	E_LightTowerState.eRed:;
		qLedGreen	:=FALSE;
		qLedYellow	:=FALSE;
		qLedRed		:=TRUE;
		qLedBlue	:=FALSE;
		IF bBuzzerMuteMemo THEN;
			eBuzzerMode:=eBuzzerOff;
		ELSE
			eBuzzerMode:=eBuzzerError;
		END_IF
		
	E_LightTowerState.eBlue:;
		qLedGreen	:=FALSE;
		qLedYellow	:=FALSE;
		qLedRed		:=FALSE;
		qLedBlue	:=TRUE;
		eBuzzerMode:=eBuzzerOff;	
				
END_CASE


IF qLedRed THEN;
	qSignal_1:=TRUE;	//wire BN
	qSignal_2:=FALSE;	//wire GY
	qSignal_3:=FALSE;	//wire BK
	qSignal_4:=FALSE;	//wire WT	
ELSIF qLedYellow THEN;
	qSignal_1:=TRUE;	//wire BN
	qSignal_2:=FALSE;	//wire GY
	qSignal_3:=FALSE;	//wire BK
	qSignal_4:=TRUE;	//wire WT	
ELSIF qLedGreen THEN;
	qSignal_1:=FALSE;	//wire BN
	qSignal_2:=FALSE;	//wire GY
	qSignal_3:=FALSE;	//wire BK
	qSignal_4:=TRUE;	//wire WT	
ELSIF qLedBlue THEN;
	qSignal_1:=FALSE;	//wire BN
	qSignal_2:=TRUE;	//wire GY
	qSignal_3:=FALSE;	//wire BK
	qSignal_4:=FALSE;	//wire WT	
ELSE;
	qSignal_1:=FALSE;	//wire BN
	qSignal_2:=FALSE;	//wire GY
	qSignal_3:=FALSE;	//wire BK
	qSignal_4:=FALSE;	//wire WT
END_IF
END_METHOD

PROPERTY pState : E_LightTowerState
GET
pState:=eLightTowerState;
END_GET
SET
eLightTowerState:=pState;
END_SET
END_PROPERTY

END_FUNCTION_BLOCK

// ---- 01 Instance/07-Mode/FB_LightTower_Control.TcPOU
FUNCTION_BLOCK FB_LightTower_Control
VAR_INPUT
	ES_State		: BOOL;
	RunProcess1		: BOOL;
	RunProcess2		: BOOL;
	RunProcess3		: BOOL;
	ModeZone1		: E_ModeZone;
	ModeZone2		: E_ModeZone;
	ModeZone3		: E_ModeZone;
END_VAR

VAR_OUTPUT
	eLightTowerState		: E_LightTowerState;
END_VAR
VAR
END_VAR

IF ES_State THEN;
	IF stOper[ModeZone1].iActOperation=E_OperationButtons.ePauseAll 
	OR stOper[ModeZone2].iActOperation=E_OperationButtons.ePauseAll
	OR stOper[ModeZone3].iActOperation=E_OperationButtons.ePauseAll
	THEN;
		eLightTowerState:= E_LightTowerState.eYellow;
	ELSIF RunProcess1 OR RunProcess2 OR RunProcess3 THEN;
		eLightTowerState:= E_LightTowerState.eGreen;
	ELSE;
		eLightTowerState:= E_LightTowerState.eBlue;
	END_IF
	
ELSE;
	eLightTowerState:= E_LightTowerState.eRed;
END_IF

END_FUNCTION_BLOCK

// ---- 03 Project/22 InterConnection/04 Mode/prg_IntCheck.TcPOU
PROGRAM prg_IntCheck
VAR_OUTPUT
	bActive_Marinade_TriB: BOOL;
	bActive_Color_TriB: BOOL;
	bActive_Marinade_Prod: BOOL;
	bActive_Color_Prod: BOOL;
END_VAR

IF fbIntCon_TriB_T1_Marin.bActive OR fbIntCon_TriB_T2_Marin.bActive THEN;
	bActive_Marinade_TriB:=TRUE;
ELSE;
	bActive_Marinade_TriB:=FALSE;
END_IF

IF fbIntCon_TriB_T3_Color.bActive OR fbIntCon_TriB_T4_Color.bActive THEN;
	bActive_Color_TriB:=TRUE;
ELSE;
	bActive_Color_TriB:=FALSE;
END_IF

IF fbIntCon_ProL_T1_Marin.bActive OR fbIntCon_ProL_T2_Marin.bActive THEN;
	bActive_Marinade_Prod:=TRUE;
ELSE;
	bActive_Marinade_Prod:=FALSE;
END_IF

IF fbIntCon_ProL_T3_Color.bActive OR fbIntCon_ProL_T4_Color.bActive THEN;
	bActive_Color_Prod:=TRUE;
ELSE;
	bActive_Color_Prod:=FALSE;
END_IF

END_PROGRAM

// ---- 00 Library/00-General/UserGroup/prg_User.TcPOU
PROGRAM prg_User
VAR
	actUser: E_userGroup:=1;
		
	ton_UserLoged: TON;
	Password: INT;
	ton_Password: TON;
	PT: BOOL;
END_VAR

ton_UserLoged(IN:=actUser<>Group1, PT:=T#10M);

IF ton_UserLoged.Q OR Password=1  THEN
	actUser:=1;
END_IF

IF Password=726 THEN
	actUser:=2;
END_IF

IF Password=345 THEN
	actUser:=3;
END_IF

IF Password=888 THEN
	actUser:=4;
END_IF


ton_Password(IN:=Password<> 0, PT:=T#1s);
IF ton_Password.Q THEN
	Password:=0;
END_IF
;

END_PROGRAM

// ---- 03 Project/22 InterConnection/00 General/prg_InterCon_Usage.TcPOU
PROGRAM prg_InterCon_Usage
VAR
END_VAR

// TriBlender  

IF fbElement[E_Element_List.eTank_1].eState_Short=E_Element_State_Short.eClean 
AND fbElement[E_Element_List.eTriBlender_Marinada].eState_Short=E_Element_State_Short.eClean
THEN;
	//eIntCon_TriB_T1_Marin:=E_InterConnection.Avalable;
END_IF

act_Call_InterConnection();

CASE eTriBlenderUsage OF
	E_TriBlenderUsage.eMarinada_T1,E_TriBlenderUsage.eMarinada_T2:;
		fbElement[E_Element_List.eTriBlender_Marinada].m_StateUpdate_Limit(value:=TRUE);		
		fbElement[E_Element_List.eTriBlender_Color].m_StateUpdate_Limit(value:=TRUE);
	
	E_TriBlenderUsage.eMarinada_Standby:;
		fbElement[E_Element_List.eTriBlender_Marinada].m_StateUpdate_Limit(value:=FALSE);
		fbElement[E_Element_List.eTriBlender_Color].m_StateUpdate_Limit(value:=TRUE);
		
	E_TriBlenderUsage.eColor_T3,E_TriBlenderUsage.eColor_T4:;	
		fbElement[E_Element_List.eTriBlender_Marinada].m_StateUpdate_Limit(value:=TRUE);		
		fbElement[E_Element_List.eTriBlender_Color].m_StateUpdate_Limit(value:=TRUE);
	
	E_TriBlenderUsage.eColor_Standby:;	
		fbElement[E_Element_List.eTriBlender_Marinada].m_StateUpdate_Limit(value:=TRUE);
		fbElement[E_Element_List.eTriBlender_Color].m_StateUpdate_Limit(value:=FALSE);
ELSE;
		fbElement[E_Element_List.eTriBlender_Marinada].m_StateUpdate_Limit(value:=FALSE);
		fbElement[E_Element_List.eTriBlender_Color].m_StateUpdate_Limit(value:=FALSE);	
END_CASE

CASE ePrL_M_Usage OF
	E_PrLine_M_LineUsage.eMarinada_T1,
	E_PrLine_M_LineUsage.eMarinada_T2:;
		fbElement[E_Element_List.eLine_Marinada].m_StateUpdate_Limit(value:=TRUE);
	E_PrLine_M_LineUsage.eNotInUse:;
		fbElement[E_Element_List.eLine_Marinada].m_StateUpdate_Limit(value:=FALSE);
END_CASE

CASE ePrL_C_Usage OF
	E_PrLine_C_Usage.eColor_T3,
	E_PrLine_C_Usage.eColor_T4:;
		fbElement[E_Element_List.eLine_Color].m_StateUpdate_Limit(value:=TRUE);
	E_PrLine_C_Usage.eNotInUse:;
		fbElement[E_Element_List.eLine_Color].m_StateUpdate_Limit(value:=FALSE);
END_CASE
(*
IF eTriBlenderPipe_In=eTriBlenderPipe_Out THEN;
	eTriBlenderPipe:=eTriBlenderPipe_In;
ELSE;
	eTriBlenderPipe:=E_TriBlenderPipe.eNone;
END_IF
*)
(*
CASE fbTriBlender_Select.eStatus OF
	E_TriBlenderSelect.eMarinade:;
		eTriBlenderPipe:=E_TriBlenderPipe.eMarinada;	
	E_TriBlenderSelect.eColor:;
		eTriBlenderPipe:=E_TriBlenderPipe.eColor;
	E_TriBlenderSelect.eDrain:;
		eTriBlenderPipe:=E_TriBlenderPipe.eNone;
ELSE;
	eTriBlenderPipe:=E_TriBlenderPipe.eNone;	
END_CASE
*)

ACTION act_Call_InterConnection:
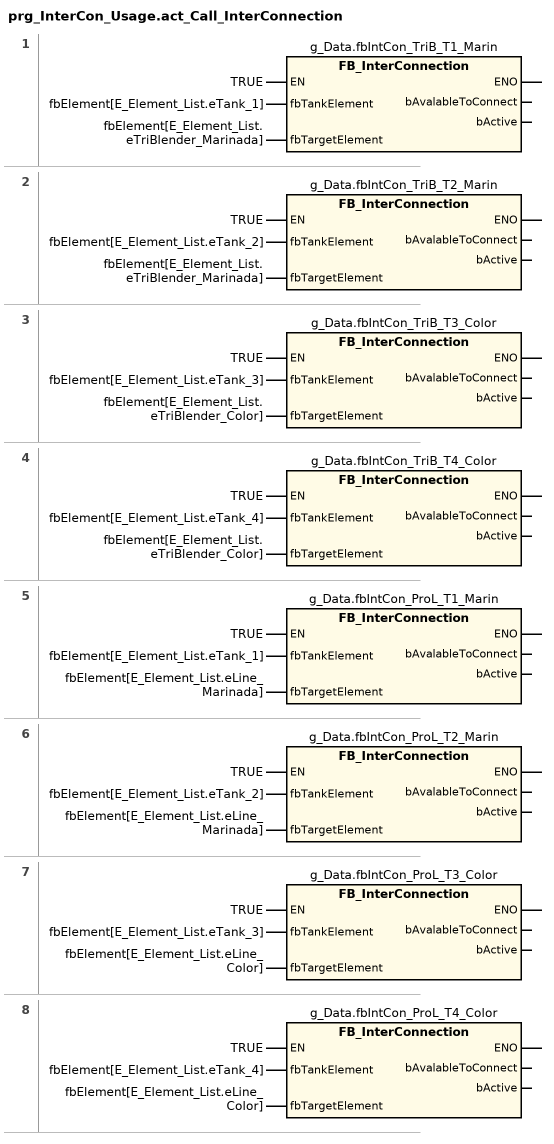
// NETWORK 1
g_Data.fbIntCon_TriB_T1_Marin(fbTankElement := fbElement[E_Element_List.eTank_1], fbTargetElement := fbElement[E_Element_List.eTriBlender_Marinada]); // FB_InterConnection

// NETWORK 2
g_Data.fbIntCon_TriB_T2_Marin(fbTankElement := fbElement[E_Element_List.eTank_2], fbTargetElement := fbElement[E_Element_List.eTriBlender_Marinada]); // FB_InterConnection

// NETWORK 3
g_Data.fbIntCon_TriB_T3_Color(fbTankElement := fbElement[E_Element_List.eTank_3], fbTargetElement := fbElement[E_Element_List.eTriBlender_Color]); // FB_InterConnection

// NETWORK 4
g_Data.fbIntCon_TriB_T4_Color(fbTankElement := fbElement[E_Element_List.eTank_4], fbTargetElement := fbElement[E_Element_List.eTriBlender_Color]); // FB_InterConnection

// NETWORK 5
g_Data.fbIntCon_ProL_T1_Marin(fbTankElement := fbElement[E_Element_List.eTank_1], fbTargetElement := fbElement[E_Element_List.eLine_Marinada]); // FB_InterConnection

// NETWORK 6
g_Data.fbIntCon_ProL_T2_Marin(fbTankElement := fbElement[E_Element_List.eTank_2], fbTargetElement := fbElement[E_Element_List.eLine_Marinada]); // FB_InterConnection

// NETWORK 7
g_Data.fbIntCon_ProL_T3_Color(fbTankElement := fbElement[E_Element_List.eTank_3], fbTargetElement := fbElement[E_Element_List.eLine_Color]); // FB_InterConnection

// NETWORK 8
g_Data.fbIntCon_ProL_T4_Color(fbTankElement := fbElement[E_Element_List.eTank_4], fbTargetElement := fbElement[E_Element_List.eLine_Color]); // FB_InterConnection
END_ACTION

END_PROGRAM

// ---- 03 Project/22 InterConnection/00 General/FB_InterConnection.TcPOU
FUNCTION_BLOCK FB_InterConnection
VAR_INPUT
	//eState_Tank		: E_Element_State_Short;
	//eState_Target	: E_Element_State_Short;
	//eProdType		: E_Product_Type;
	//eTargetTape		: E_Element_Type:=E_Element_Type.eNotSelected;
	reqConnect: BOOL;
	reqDisconnect: BOOL;

END_VAR
VAR_OUTPUT
	bAvalableToConnect: BOOL;
	bAvalableToDisconnect: BOOL;
	bActive: BOOL;
END_VAR
VAR



END_VAR

VAR_IN_OUT
	fbTankElement: FB_Element;
	fbTargetElement: FB_Element;	
END_VAR

act_Avalable();
act_Active();




IF reqConnect THEN;
	m_Connect();
	reqConnect:=FALSE;
END_IF

IF reqDisconnect THEN;
	m_Disconnect();
	reqDisconnect:=FALSE;
END_IF

IF fbTankElement.eInterConnect <> E_InterConnection.NotConnected 
OR fbTargetElement.eInterConnect <> E_InterConnection.NotConnected
THEN;
	m_At_Connected_Pause();
	m_At_Connected_Play();
END_IF

ACTION act_Active:
//fbTargetElement.eState_Long:=fbTankElement.eState_Long;
IF bActive THEN;
	fbTargetElement.m_InterConnected_State(eState_Long_Set:=fbTankElement.eState_Long);
	//fbTargetElement.ExpirationTime:=fbTankElement.ExpirationTime;
	
	CASE fbTargetElement.eType OF		
		E_Element_Type.eLine:;
			//fbTankElement.m_InterConnect(value:=E_InterConnection.ConnToLine);			
		E_Element_Type.eTriBlender:;
			//fbTankElement.m_InterConnect(value:=E_InterConnection.ConnToTriBlender);		
	END_CASE
	//fbTargetElement.m_InterConnect(value:=E_InterConnection.ConnToTank);
	
	CASE fbTankElement.eState_Short OF
		E_Element_State_Short.eNotClean,
		E_Element_State_Short.eClean:;
				//fbTargetElement.ExpirationMode:=E_ExTime.eCIP;

		E_Element_State_Short.eProduct:;
				//fbTargetElement.ExpirationMode:=E_ExTime.eLine;
	END_CASE	

ELSE;
	//fbTankElement.m_Disconnect();
	//fbTargetElement.m_Disconnect();
END_IF
END_ACTION

ACTION act_At_Connected_Pause:

/// Master case
IF fbTankElement.m_Get_Oper_Pause_Puls() THEN;
	CASE fbTankElement.eInterConnect OF 
		E_InterConnection.NotConnected:;
		E_InterConnection.ConnToCIP:;
				// set pause to CIP
				stOper[E_ModeZone.eCIP].bSetPause:=TRUE;
				
		E_InterConnection.ConnToTank:;
				//Not avilble 
		E_InterConnection.ConnToLine:;
				IF fbTargetElement.m_Get_Type()=E_Element_Type.eLine THEN;
					fbTargetElement.m_Set_Oper_Pause();
				END_IF
		E_InterConnection.ConnToTriBlender:;
				IF fbTargetElement.m_Get_Type()=E_Element_Type.eTriBlender THEN;
					fbTargetElement.m_Set_Oper_Pause();
				END_IF				
	END_CASE	
END_IF


/// Slave case
IF fbTargetElement.m_Get_Oper_Pause_Puls() THEN;
	CASE fbTargetElement.eInterConnect OF 
		E_InterConnection.NotConnected:;
		E_InterConnection.ConnToCIP:;
				// set pause to CIP
				stOper[E_ModeZone.eCIP].bSetPause:=TRUE;
				
		E_InterConnection.ConnToTank:;
				IF TRUE
				AND fbTargetElement.m_Get_Type()=E_Element_Type.eLine
				AND fbTankElement.eInterConnect=E_InterConnection.ConnToLine THEN;
					fbTankElement.m_Set_Oper_Pause();
				END_IF
				
				IF TRUE
				AND fbTargetElement.m_Get_Type()=E_Element_Type.eTriBlender
				AND fbTankElement.eInterConnect=E_InterConnection.ConnToTriBlender THEN;
					fbTankElement.m_Set_Oper_Pause();
				END_IF
								
		E_InterConnection.ConnToLine:;
				//Not avilble 
		E_InterConnection.ConnToTriBlender:;
				//Not avilble 			
	END_CASE	
END_IF

// CIP Case
IF stOper[E_ModeZone.eCIP].b_rt_Pause 
AND	fbTankElement.eInterConnect=E_InterConnection.ConnToCIP
THEN;	
	fbTankElement.m_Set_Oper_Pause();
END_IF

IF stOper[E_ModeZone.eCIP].b_rt_Pause 
AND	fbTargetElement.eInterConnect=E_InterConnection.ConnToCIP
THEN;	
	fbTargetElement.m_Set_Oper_Pause();
END_IF
END_ACTION

ACTION act_At_Connected_Play:

/// Master case
IF fbTankElement.m_Get_Oper_Play_Puls() THEN;
	CASE fbTankElement.eInterConnect OF 
		E_InterConnection.NotConnected:;
		E_InterConnection.ConnToCIP:;
				// set Play to CIP
				//stOper[E_ModeZone.eCIP].bSetPlay:=TRUE;
				
		E_InterConnection.ConnToTank:;
				//Not avilble 
		E_InterConnection.ConnToLine:;
				IF fbTargetElement.m_Get_Type()=E_Element_Type.eLine THEN;
					fbTargetElement.m_Set_Oper_Play();
				END_IF
		E_InterConnection.ConnToTriBlender:;
				IF fbTargetElement.m_Get_Type()=E_Element_Type.eTriBlender THEN;
					fbTargetElement.m_Set_Oper_Play();
				END_IF				
	END_CASE	
END_IF


// CIP Case
IF stOper[E_ModeZone.eCIP].b_rt_Play 
AND	fbTankElement.eInterConnect=E_InterConnection.ConnToCIP
THEN;	
	fbTankElement.m_Set_Oper_Play();
END_IF

IF stOper[E_ModeZone.eCIP].b_rt_Play 
AND	fbTargetElement.eInterConnect=E_InterConnection.ConnToCIP
THEN;	
	fbTargetElement.m_Set_Oper_Play();
END_IF
END_ACTION

ACTION act_Avalable:
// To Connect
CASE fbTargetElement.eType OF
	E_Element_Type.eTriBlender:;
			IF (eTriBlenderUsage=E_TriBlenderUsage.eNotInUse 
			OR(eTriBlenderUsage=E_TriBlenderUsage.eMarinada_Standby 
				AND fbTankElement.eProdType=E_Product_Type.Marinada)
			OR(eTriBlenderUsage=E_TriBlenderUsage.eColor_Standby 
				AND fbTankElement.eProdType=E_Product_Type.Color))
			//AND fbElement[E_Element_List.eTriBlender_Marinada].eState_Short<>E_Element_State_Short.eNotClean	
			//AND fbElement[E_Element_List.eTriBlender_Color].eState_Short<>E_Element_State_Short.eNotClean
			AND fbTankElement.eInterConnect=E_InterConnection.NotConnected	
			AND fbTargetElement.eInterConnect=E_InterConnection.NotConnected	
			
			// Pipe check
			(*AND ((fbTargetElement.eProdType=E_Product_Type.Marinada AND eTriBlenderPipe=E_TriBlenderPipe.eMarinada)
							OR
				(fbTargetElement.eProdType=E_Product_Type.Color AND eTriBlenderPipe=E_TriBlenderPipe.eColor))*)
		
			THEN;
				IF (fbTankElement.eState_Short=E_Element_State_Short.eClean 
					OR fbTankElement.eState_Short=E_Element_State_Short.eProduct
					)
				AND (fbTargetElement.eState_Short=E_Element_State_Short.eClean 
					OR fbTargetElement.eState_Short=E_Element_State_Short.eProduct)
				THEN;
					bAvalableToConnect:=TRUE;
				ELSE;
					bAvalableToConnect:=FALSE;
				END_IF	
			ELSE;
				bAvalableToConnect:=FALSE;
			END_IF
		
			IF eTriBlenderUsage=E_TriBlenderUsage.eMarinada_Standby
			AND fbTargetElement.eProdType=E_Product_Type.Marinada
			AND	fbTargetElement.eState_Short=E_Element_State_Short.eClean
			THEN;
				eTriBlenderUsage:=E_TriBlenderUsage.eNotInUse;
			END_IF

			IF eTriBlenderUsage=E_TriBlenderUsage.eColor_Standby
			AND fbTargetElement.eProdType=E_Product_Type.Color
			AND	fbTargetElement.eState_Short=E_Element_State_Short.eClean
			THEN;
				eTriBlenderUsage:=E_TriBlenderUsage.eNotInUse;
			END_IF
			
	
	E_Element_Type.eLine:;
	
			IF ((fbTankElement.eProdType=E_Product_Type.Marinada
				AND ePrL_M_Usage=E_PrLine_M_LineUsage.eNotInUse) 
			OR(fbTankElement.eProdType=E_Product_Type.Color
				AND ePrL_C_Usage=E_PrLine_C_Usage.eNotInUse)) 
			AND fbTankElement.eInterConnect=E_InterConnection.NotConnected
			AND fbTargetElement.eInterConnect=E_InterConnection.NotConnected 
			THEN;
				IF (fbTankElement.eState_Short=E_Element_State_Short.eProduct 
					//OR fbTankElement.eState_Short=E_Element_State_Short.eClean)
					)
				AND (fbTargetElement.eState_Short=E_Element_State_Short.eProduct 
					OR fbTargetElement.eState_Short=E_Element_State_Short.eClean)
				THEN;
					bAvalableToConnect:=TRUE;
				ELSE;
					bAvalableToConnect:=FALSE;
				END_IF			
			ELSE;
				bAvalableToConnect:=FALSE;
			END_IF
	
END_CASE

// To Disconnect
CASE fbTargetElement.eType OF
	E_Element_Type.eTriBlender:;
		IF bActive THEN;// AND fbTankElement.eState_Long<>E_Element_State_Long.eProduction
			bAvalableToDisconnect:=TRUE;
		ELSE;
			bAvalableToDisconnect:=FALSE;
		END_IF
	E_Element_Type.eLine:;
		IF bActive AND (fbTankElement.eState_Long=E_Element_State_Long.eProduction 
						OR fbTankElement.eState_Long_Expiered=E_Element_State_Long.eProduction)
		THEN;
			bAvalableToDisconnect:=TRUE;
		ELSE;
			bAvalableToDisconnect:=FALSE;
		END_IF	
END_CASE
END_ACTION

METHOD m_At_Connected_Pause : BOOL
VAR_INPUT
END_VAR

/// Master case
IF fbTankElement.m_Get_Oper_Pause_Puls() THEN;
	CASE fbTankElement.eInterConnect OF 
		E_InterConnection.NotConnected:;
		E_InterConnection.ConnToCIP:;
				// set pause to CIP
				stOper[E_ModeZone.eCIP].bSetPause:=TRUE;
				RETURN;
		E_InterConnection.ConnToTank:;
				//Not avilble 
		E_InterConnection.ConnToLine:;
				IF fbTargetElement.m_Get_Type()=E_Element_Type.eLine THEN;
					fbTargetElement.m_Set_Oper_Pause();
					RETURN;
				END_IF
		E_InterConnection.ConnToTriBlender:;
				IF fbTargetElement.m_Get_Type()=E_Element_Type.eTriBlender THEN;
					fbTargetElement.m_Set_Oper_Pause();
					RETURN;
				END_IF				
	END_CASE	
END_IF


/// Slave case
IF fbTargetElement.m_Get_Oper_Pause_Puls() THEN;
	CASE fbTargetElement.eInterConnect OF 
		E_InterConnection.NotConnected:;
		E_InterConnection.ConnToCIP:;
				// set pause to CIP
				stOper[E_ModeZone.eCIP].bSetPause:=TRUE;
				RETURN;
		E_InterConnection.ConnToTank:;
				IF TRUE
				AND fbTargetElement.m_Get_Type()=E_Element_Type.eLine
				AND fbTankElement.eInterConnect=E_InterConnection.ConnToLine THEN;
					fbTankElement.m_Set_Oper_Pause();
					RETURN;
				END_IF
				
				IF TRUE
				AND fbTargetElement.m_Get_Type()=E_Element_Type.eTriBlender
				AND fbTankElement.eInterConnect=E_InterConnection.ConnToTriBlender THEN;
					fbTankElement.m_Set_Oper_Pause();
					RETURN;
				END_IF
								
		E_InterConnection.ConnToLine:;
				//Not avilble 
		E_InterConnection.ConnToTriBlender:;
				//Not avilble 			
	END_CASE	
END_IF

// CIP Case
IF stOper[E_ModeZone.eCIP].b_rt_Pause 
AND	fbTankElement.eInterConnect=E_InterConnection.ConnToCIP
THEN;	
	fbTankElement.m_Set_Oper_Pause();
	RETURN;
END_IF

IF stOper[E_ModeZone.eCIP].b_rt_Pause 
AND	fbTargetElement.eInterConnect=E_InterConnection.ConnToCIP
THEN;	
	fbTargetElement.m_Set_Oper_Pause();
	RETURN;
END_IF
END_METHOD

METHOD m_At_Connected_Play : BOOL
VAR_INPUT
END_VAR

/// Master case
IF fbTankElement.m_Get_Oper_Play_Puls() THEN;
	CASE fbTankElement.eInterConnect OF 
		E_InterConnection.NotConnected:;
		E_InterConnection.ConnToCIP:;
				// Not avilble				
		E_InterConnection.ConnToTank:;
				//Not avilble 
		E_InterConnection.ConnToLine:;
				IF fbTargetElement.m_Get_Type()=E_Element_Type.eLine THEN;
					fbTargetElement.m_Set_Oper_Play();
					RETURN;
				END_IF
		E_InterConnection.ConnToTriBlender:;
				IF fbTargetElement.m_Get_Type()=E_Element_Type.eTriBlender THEN;
					fbTargetElement.m_Set_Oper_Play();
					RETURN;
				END_IF				
	END_CASE	
END_IF


// CIP Case
IF stOper[E_ModeZone.eCIP].b_rt_Play 
AND	fbTankElement.eInterConnect=E_InterConnection.ConnToCIP
THEN;	
	fbTankElement.m_Set_Oper_Play();
	RETURN;
END_IF

IF stOper[E_ModeZone.eCIP].b_rt_Play 
AND	fbTargetElement.eInterConnect=E_InterConnection.ConnToCIP
THEN;	
	fbTargetElement.m_Set_Oper_Play();
	RETURN;
END_IF
END_METHOD

METHOD m_Connect : BOOL
VAR_INPUT
END_VAR
IF bAvalableToConnect THEN;
	
	CASE fbTankElement.eElementID OF
		E_Element_List.eTank_1:;
				CASE fbTargetElement.eElementID OF
					E_Element_List.eTriBlender_Marinada:;
						eTriBlenderUsage:=E_TriBlenderUsage.eMarinada_T1;
						fbTankElement.m_InterConnect(value:=E_InterConnection.ConnToTriBlender);
					E_Element_List.eLine_Marinada:;
						ePrL_M_Usage:=E_PrLine_M_LineUsage.eMarinada_T1;
						fbTankElement.m_InterConnect(value:=E_InterConnection.ConnToLine);
				END_CASE								
				
		E_Element_List.eTank_2:;		
				CASE fbTargetElement.eElementID OF
					E_Element_List.eTriBlender_Marinada:;
						eTriBlenderUsage:=E_TriBlenderUsage.eMarinada_T2;
						fbTankElement.m_InterConnect(value:=E_InterConnection.ConnToTriBlender);
					E_Element_List.eLine_Marinada:;
						ePrL_M_Usage:=E_PrLine_M_LineUsage.eMarinada_T2;
						fbTankElement.m_InterConnect(value:=E_InterConnection.ConnToLine);
				END_CASE		
		
				
		E_Element_List.eTank_3:;
				CASE fbTargetElement.eElementID OF
					E_Element_List.eTriBlender_Color:;
						eTriBlenderUsage:=E_TriBlenderUsage.eColor_T3;
						fbTankElement.m_InterConnect(value:=E_InterConnection.ConnToTriBlender);
					E_Element_List.eLine_Color:;
						ePrL_C_Usage:=E_PrLine_C_Usage.eColor_T3;
						fbTankElement.m_InterConnect(value:=E_InterConnection.ConnToLine);
				END_CASE
						
		E_Element_List.eTank_4:;
				CASE fbTargetElement.eElementID OF
					E_Element_List.eTriBlender_Color:;
						eTriBlenderUsage:=E_TriBlenderUsage.eColor_T4;
						fbTankElement.m_InterConnect(value:=E_InterConnection.ConnToTriBlender);
					E_Element_List.eLine_Color:;
						ePrL_C_Usage:=E_PrLine_C_Usage.eColor_T4;
						fbTankElement.m_InterConnect(value:=E_InterConnection.ConnToLine);
				END_CASE		
						
	END_CASE
	fbTargetElement.m_InterConnect(value:=E_InterConnection.ConnToTank);
	bActive:=TRUE;
ELSE;

END_IF
END_METHOD

METHOD m_Disconnect : BOOL
VAR_INPUT
END_VAR
IF bActive AND fbTankElement.eState_Long<>E_Element_State_Long.eProduction THEN;
	IF fbTargetElement.eType=E_Element_Type.eTriBlender THEN;
		IF fbTargetElement.eState_Short=E_Element_State_Short.eProduct THEN;
			IF fbTankElement.eProdType=E_Product_Type.Marinada 
			AND fbTargetElement.memoDissolving_active
			THEN;
				eTriBlenderUsage:=E_TriBlenderUsage.eMarinada_Standby;
			END_IF
			IF fbTankElement.eProdType=E_Product_Type.Color 
			AND fbTargetElement.memoDissolving_active
			THEN;
				eTriBlenderUsage:=E_TriBlenderUsage.eColor_Standby;
			END_IF
		ELSE;
			eTriBlenderUsage:=E_TriBlenderUsage.eNotInUse;
		END_IF
		
		
	ELSIF fbTargetElement.eType=E_Element_Type.eLine THEN;
		IF fbTankElement.eProdType=E_Product_Type.Marinada THEN;
			ePrL_M_Usage:=E_PrLine_M_LineUsage.eNotInUse;
		END_IF
		IF fbTankElement.eProdType=E_Product_Type.Color THEN;
			ePrL_C_Usage:=E_PrLine_C_Usage.eNotInUse;
		END_IF		
	END_IF
	
	fbTankElement.m_Disconnect();
	fbTargetElement.m_Disconnect();
	
	IF fbTankElement.ExpirationTime<T#2H THEN;
		//fbTargetElement.ExpirationTime:=T#1H;
	ELSE;
		//fbTargetElement.ExpirationTime:=T#2h;
	END_IF
	
	bActive:=FALSE;
END_IF
END_METHOD

END_FUNCTION_BLOCK

// ---- 03 Project/10 Element/FB_Element.TcPOU
FUNCTION_BLOCK FB_Element// EXTENDS FB_SFC_Cycle IMPLEMENTS ITF_FB_SFC_Cycle
VAR_INPUT
	eElementID			: E_Element_List;

END_VAR
VAR_OUTPUT
	event_StateUpdate	: INT; // for HMI
END_VAR



VAR
	eType				: E_Element_Type;
	eProdType			: E_Product_Type;
	eState_Long			: E_Element_State_Long;
	eState_Short		: E_Element_State_Short;
	eState_Long_last	: E_Element_State_Long;
	eState_Long_Expiered: E_Element_State_Long;





	i: INT;
	sState_Time			: STRING;
	sTimeToExpiration	: STRING;
	tTimeToExpiration	: TIME;
	tStateTime			: TIME;

	
	sElementID			: STRING;
	eInterConnect		: E_InterConnection;
	memoDissolving_active		: BOOL;
	bStateUpdate_Limited		: BOOL;

	stCIP_Request		: ST_CIP_Request;
	stCIP_RequestActive	: ST_CIP_Request;

	bTakePosInCIPBuffer_Partial		: BOOL;
	bTakePosInCIPBuffer_Full		: BOOL;
	bTakePosInCIPBuffer_Detergent	: BOOL;
	bError: BOOL;	
	
	eProdStatus			: E_Prod_Status;
	eFilling_State		: E_Filling_State;
	
	fbEvent_echo: FB_Event_echo;

END_VAR

VAR PERSISTENT
	tsStateChange				: TimeStruct;
	tsCIP						: TimeStruct;
	tsWater						: TimeStruct;
	tsProduction				: TimeStruct;
	tsProductionLine			: TimeStruct;
	tsProductionLineStby		: TimeStruct;
	
	
	tExpirationTime				: TIME:=T#48H;
	ExDuration_Product			: TIME:=T#48H; 	//Expiration from loaded ricipe
	ExDuration_Water			: TIME:=T#48H; 	//Expiration from loaded ricipe
	
	eExTime						: E_ExTime;


END_VAR


VAR_IN_OUT
	stOperation		: ST_OperationButtons;	
END_VAR

i:=i+1;
//m_Set_SFCFlags_Reference();
//SUPER^();
fbEvent_echo(echo=>event_StateUpdate);
act_StateMachine();
act_StateChange_WatchGog();

sElementID:=TO_STRING(eElementID);

CASE eType OF 
	E_Element_Type.eTank:;
				act_Tank();
	E_Element_Type.eTriBlender:;
				act_TriBlender();
	E_Element_Type.eLine:;
				act_Line();

END_CASE

CASE eElementID OF
	E_Element_List.eTank_1:;
				eType:=E_Element_Type.eTank;
				eProdType:=E_Product_Type.Marinada;
				stCIP_Request.eClient:=E_CIP_Usage.eTank_1;
	E_Element_List.eTank_2:;
				eType:=E_Element_Type.eTank;
				eProdType:=E_Product_Type.Marinada;
				stCIP_Request.eClient:=E_CIP_Usage.eTank_2;
	E_Element_List.eTank_3:;
				eType:=E_Element_Type.eTank;
				eProdType:=E_Product_Type.Color;
				stCIP_Request.eClient:=E_CIP_Usage.eTank_3;
	E_Element_List.eTank_4:;
				eType:=E_Element_Type.eTank;
				eProdType:=E_Product_Type.Color;
				stCIP_Request.eClient:=E_CIP_Usage.eTank_4;
	E_Element_List.eTriBlender_Marinada:;
				eType:=E_Element_Type.eTriBlender;
				eProdType:=E_Product_Type.Marinada;		
				stCIP_Request.eClient:=E_CIP_Usage.eTriBlender_Marinada;
	E_Element_List.eTriBlender_Color:;
				eType:=E_Element_Type.eTriBlender;
				eProdType:=E_Product_Type.Color;
				stCIP_Request.eClient:=E_CIP_Usage.eTriBlender_Color;
	E_Element_List.eLine_Marinada:;
				eType:=E_Element_Type.eLine;
				eProdType:=E_Product_Type.Marinada;
				stCIP_Request.eClient:=E_CIP_Usage.eLine_Marinada;
	E_Element_List.eLine_Color:;
				eType:=E_Element_Type.eLine;
				eProdType:=E_Product_Type.Color;
				stCIP_Request.eClient:=E_CIP_Usage.eLine_Color;
END_CASE


IF bTakePosInCIPBuffer_Partial THEN;
	stCIP_Request.eType:=E_CIP_Type.R_Water;
	fbCIP.m_TakePosInCIPBuffer(stCIP_Request:=stCIP_Request);
	bTakePosInCIPBuffer_Partial:=FALSE;
END_IF

IF bTakePosInCIPBuffer_Detergent THEN;
	stCIP_Request.eType:=E_CIP_Type.Detergent;
	fbCIP.m_TakePosInCIPBuffer(stCIP_Request:=stCIP_Request);
	bTakePosInCIPBuffer_Detergent:=FALSE;
END_IF

IF bTakePosInCIPBuffer_Full THEN;
	stCIP_Request.eType:=E_CIP_Type.Full;
	fbCIP.m_TakePosInCIPBuffer(stCIP_Request:=stCIP_Request);
	bTakePosInCIPBuffer_Full:=FALSE;
END_IF

stCIP_RequestActive.eType:=E_CIP_Type.NotSelected;
FOR i:=0 TO 9 DO
	IF arCIP_RequestBufer[i].eClient=stCIP_Request.eClient
	AND arCIP_RequestBufer[i].eType>stCIP_RequestActive.eType THEN;
		stCIP_RequestActive.eType:=arCIP_RequestBufer[i].eType;
	END_IF
END_FOR

m_TimeToExpiration();

ACTION act_Line:

END_ACTION

ACTION act_StateChange_WatchGog:
IF eState_Long<>eState_Long_last THEN;
	IF eState_Long=E_Element_State_Long.eExpired THEN;
		eState_Long_Expiered:=eState_Long_last;
	ELSE;
		eState_Long_Expiered:=E_Element_State_Long.eOff;
	END_IF

	IF eState_Long=E_Element_State_Long.eWaterReady THEN;
		IF  eState_Long_last=E_Element_State_Long.eCIP_5_Done THEN;
			//tsWater:=stSystemTime;
			m_Set_TimeToExpirationMode(eExTime_set:=E_ExTime.eWater);
		ELSE;
			// do nothing here...
		END_IF
		
	ELSIF eState_Long>=E_Element_State_Long.eReady THEN;
		IF eState_Long=E_Element_State_Long.eReady
		AND NOT memoDissolving_active THEN; // state updated manualy
			m_Set_Dissolveng_active_memo();
		ELSE; // state update during dissolving status
			// do nothing here...
		END_IF
	ELSE;
		//tsCIP:=stSystemTime;
		m_Set_TimeToExpirationMode(eExTime_set:=E_ExTime.eCIP);
		
	END_IF
	
	eState_Long_last:=eState_Long;
	
	fbEvent_echo.event(); // for HMI
END_IF

tStateTime:=TO_TIME(SYSTEMTIME_TO_DT(stSystemTime)-SYSTEMTIME_TO_DT(tsStateChange));

sState_Time:=prg_RealClock.m_DeltaTime(stStartTime:=tsStateChange);
sTimeToExpiration:=prg_RealClock.mTime_to_String_HMI(tInputTime:=tTimeToExpiration, iSecondDisplay:=TRUE);

sState_Time:= CONCAT(sState_Time, '(');
sState_Time:= CONCAT(sState_Time, sTimeToExpiration);
sState_Time:= CONCAT(sState_Time, ')');

CASE eExTime OF 
	E_ExTime.eCIP:sState_Time:= CONCAT(sState_Time, '/C');
	E_ExTime.eLine:sState_Time:= CONCAT(sState_Time, '/L');
	E_ExTime.eLineStby:sState_Time:= CONCAT(sState_Time, '/LS');
	E_ExTime.eProduct:sState_Time:= CONCAT(sState_Time, '/P');
	E_ExTime.eWater:sState_Time:= CONCAT(sState_Time, '/W');
	
END_CASE
END_ACTION

ACTION act_StateMachine:
CASE eState_Long OF
	E_Element_State_Long.eOff,
	E_Element_State_Long.eStandby,
	E_Element_State_Long.eNotClean,
	E_Element_State_Long.eCIP_1_Rinzed,
	E_Element_State_Long.eCIP_2_Deterged,
	E_Element_State_Long.eCIP_3_Deterged_Clean,	
	E_Element_State_Long.eCIP_4_Sanitized:;
				eState_Short:=E_Element_State_Short.eNotClean;
					ExpirationTime:=ExDuration_Default;
	E_Element_State_Long.eCIP_5_Done:;
				eState_Short:=E_Element_State_Short.eClean;
					memoDissolving_active:=FALSE;
	E_Element_State_Long.eWaterReady:;	
				IF memoDissolving_active THEN;
					eState_Short:=E_Element_State_Short.eProduct;
				ELSE;
					eState_Short:=E_Element_State_Short.eClean;
				END_IF
	E_Element_State_Long.eReady,
	E_Element_State_Long.eProduction,
	E_Element_State_Long.eEmpty:;	
				eState_Short:=E_Element_State_Short.eProduct;
	E_Element_State_Long.eExpired:;
				//
	
END_CASE
END_ACTION

ACTION act_Tank:
;
END_ACTION

ACTION act_TriBlender:
(*
IF eInterConnect=E_InterConnection.ConnToCIP 
AND eElementID=E_Element_List.eTriBlender_Marinada
AND eTriBlenderPipe<>E_TriBlenderPipe.eMarinada
THEN;
	bError:=TRUE;
ELSE;
	bError:=FALSE;
END_IF
*)
END_ACTION

PROPERTY ExpirationMode : E_ExTime
GET
ExpirationMode:=eExTime;
END_GET
SET
eExTime:=ExpirationMode;
END_SET
END_PROPERTY

PROPERTY ExpirationTime : TIME
GET
ExpirationTime:=tExpirationTime;
END_GET
SET
tExpirationTime:=ExpirationTime;
END_SET
END_PROPERTY

PROPERTY Interconnect : E_InterConnection
GET
Interconnect:=m_Get_InterConnection();
END_GET
SET
END_SET
END_PROPERTY

METHOD m_Disconnect : BOOL
VAR_INPUT
END_VAR
eInterConnect:=E_InterConnection.NotConnected;
CASE eType OF
	E_Element_Type.eTank:;					
			//
	E_Element_Type.eTriBlender,
	E_Element_Type.eLine:;
			//tsProductionLineStby:=stSystemTime;
			m_Set_TimeToExpirationMode(eExTime_set:=E_ExTime.eLineStby);
END_CASE
END_METHOD

METHOD m_Get_CIP_Avilable : BOOL
VAR_INPUT
END_VAR
IF TRUE 
AND (eInterConnect=E_InterConnection.NotConnected OR eInterConnect=E_InterConnection.ConnToCIP)
AND TRUE
THEN;
	m_Get_CIP_Avilable:=TRUE;
ELSE;
	m_Get_CIP_Avilable:=FALSE;
END_IF
END_METHOD

METHOD m_Get_InterConnection : E_InterConnection
VAR_INPUT
END_VAR

m_Get_InterConnection:=eInterConnect;
END_METHOD

METHOD m_Get_Oper_Pause_Puls : BOOL
VAR_INPUT
END_VAR
m_Get_Oper_Pause_Puls:=stOperation.b_rt_Pause;
END_METHOD

METHOD m_Get_Oper_Pause_State : BOOL
VAR_INPUT
END_VAR
IF stOperation.b_rt_Pause THEN;
	m_Get_Oper_Pause_State:=TRUE;
ELSE;
	m_Get_Oper_Pause_State:=FALSE;
END_IF
END_METHOD

METHOD m_Get_Oper_Play_Puls : BOOL
VAR_INPUT
END_VAR
m_Get_Oper_Play_Puls:=stOperation.b_rt_Play;
END_METHOD

METHOD m_Get_Oper_Play_State : BOOL
VAR_INPUT
END_VAR
IF stOperation.iActOperation=E_OperationButtons.ePlayAll THEN;
	m_Get_Oper_Play_State:=TRUE;
ELSE;
	m_Get_Oper_Play_State:=FALSE;
END_IF
END_METHOD

METHOD m_Get_State : E_Element_State_Long
VAR_INPUT
END_VAR
m_Get_State:=eState_Long;
END_METHOD

METHOD m_Get_State_Short : E_Element_State_Short
VAR_INPUT
END_VAR
m_Get_State_Short:=eState_Short;
END_METHOD

METHOD m_Get_TimeToExpirationMode : TIME
VAR_INPUT
	eExTime_check		: E_ExTime;
END_VAR

VAR
	tsStateChange_local				: TimeStruct;
	tModeTime		: TIME;
	tModeDuration	: TIME;

END_VAR
CASE eExTime_check OF
	E_ExTime.eCIP:;
			tsStateChange_local:=tsCIP;
			tModeDuration:=ExDuration_Default;
	E_ExTime.eWater:;
			tsStateChange_local:=tsWater;
			tModeDuration:=ExDuration_Water;
	E_ExTime.eProduct:;
			tsStateChange_local:=tsProduction;	
			tModeDuration:=ExDuration_Product;
	E_ExTime.eLine :;
			tsStateChange_local:=tsProductionLine;
			tModeDuration:=ExDuration_Default_Line;
	E_ExTime.eLineStby:;
			tsStateChange_local:=tsProductionLineStby;
			tModeDuration:=ExDuration_Default_LineStandby;
END_CASE
tModeTime:=TO_TIME(SYSTEMTIME_TO_DT(stSystemTime)-SYSTEMTIME_TO_DT(tsStateChange_local));
m_Get_TimeToExpirationMode:=tModeDuration-tModeTime;
END_METHOD

METHOD m_Get_Type : E_Element_Type
VAR_INPUT
END_VAR
m_Get_Type:=eType;
END_METHOD

METHOD m_InterConnect : BOOL
VAR_INPUT
	value: E_InterConnection;
END_VAR
IF eInterConnect=E_InterConnection.NotConnected 
OR eInterConnect=value
THEN;
	eInterConnect:=value;
	m_InterConnect:=TRUE;
ELSE;
	m_InterConnect:=FALSE;
END_IF
END_METHOD

METHOD m_InterConnected_State : BOOL
VAR_INPUT
	eState_Long_Set			: E_Element_State_Long;
END_VAR

IF (eState_Long_Set>eState_Long 
OR eState_Long_Set=E_Element_State_Long.eNotClean)
AND eState_Long_Set<=E_Element_State_Long.eProduction
THEN;
	eState_Long:=eState_Long_Set;
END_IF
END_METHOD

METHOD m_Set_Dissolveng_active_memo : BOOL
VAR_INPUT
END_VAR
IF NOT memoDissolving_active THEN;
	
	
	IF eInterConnect=E_InterConnection.ConnToTank THEN;
		//tsProductionLine:=stSystemTime;
		m_Set_TimeToExpirationMode(eExTime_set:=E_ExTime.eLine);
	ELSE; //element is production tank
		//tsProduction:=stSystemTime;
		m_Set_TimeToExpirationMode(eExTime_set:=E_ExTime.eProduct);
	END_IF
	
END_IF
memoDissolving_active:=TRUE;
fbEvent_echo.event();
END_METHOD

METHOD m_Set_ExpirationDuration : BOOL
VAR_INPUT
	eExTime_set		: E_ExTime;
	setTime			: TIME;

END_VAR
CASE eExTime_set OF
	E_ExTime.eCIP:;
			
	E_ExTime.eWater:;
			ExDuration_Water:=setTime;
			m_Set_ExpirationDuration:=TRUE;
	E_ExTime.eProduct:;
			ExDuration_Product:=setTime;	
			m_Set_ExpirationDuration:=TRUE;
	E_ExTime.eLine :;
			
	E_ExTime.eLineStby:;
			
END_CASE
END_METHOD

METHOD m_Set_Oper_Pause
VAR_INPUT
END_VAR
IF stOperation.iActOperation<>E_OperationButtons.ePauseAll THEN;
	stOperation.bSetPause:=TRUE;
END_IF
END_METHOD

METHOD m_Set_Oper_Play
VAR_INPUT
END_VAR
IF stOperation.iActOperation<>E_OperationButtons.ePlayAll THEN;
	stOperation.bSetPlay:=TRUE;
END_IF
END_METHOD

METHOD m_Set_SFCFlags_Reference : BOOL
//Set reference to SFC flags

refSFC.SFCInit REF= SFCInit;
refSFC.SFCReset REF= SFCReset;
refSFC.SFCError REF= SFCError;
refSFC.SFCEnableLimit REF= SFCEnableLimit;
refSFC.SFCErrorStep REF= SFCErrorStep;
refSFC.SFCErrorPOU REF= SFCErrorPOU;
refSFC.SFCQuitError REF= SFCQuitError;
refSFC.SFCPause REF= SFCPause;
refSFC.SFCTrans REF= SFCTrans;
refSFC.SFCCurrentStep REF= SFCCurrentStep;
refSFC.SFCTip REF= SFCTip;
refSFC.SFCTipMode REF= SFCTipMode;

// Cycle handle for SFC
m_SFC_Handle();
END_METHOD

METHOD m_Set_State : BOOL
VAR_INPUT
	eState_Long_Set			: E_Element_State_Long;
END_VAR
(*
IF eState_Long_Set>eState_Long 
OR eState_Long_Set=E_Element_State_Long.eNotClean
THEN;
	eState_Long:=eState_Long_Set;
END_IF
*)
eState_Long:=eState_Long_Set;
END_METHOD

METHOD m_Set_TimeToExpirationMode : TIME
VAR_INPUT
	eExTime_set		: E_ExTime;
END_VAR

VAR
	tsSet				: TimeStruct;
	tsStateChange_local				: TimeStruct;
	tModeTime		: TIME;
	tModeDuration	: TIME;

END_VAR
tsSet:=stSystemTime;
CASE eExTime_set OF
	E_ExTime.eCIP:;
			tsStateChange_local:=tsCIP:=tsSet;
			tModeDuration:=ExDuration_Default;
	E_ExTime.eWater:;
			tsStateChange_local:=tsWater:=tsSet;
			tModeDuration:=ExDuration_Water;
	E_ExTime.eProduct:;
			tsStateChange_local:=tsProduction:=tsSet;	
			tModeDuration:=ExDuration_Product;
	E_ExTime.eLine :;
			tsStateChange_local:=tsProductionLine:=tsSet;
			tModeDuration:=ExDuration_Default_Line;
	E_ExTime.eLineStby:;
			tsStateChange_local:=tsProductionLineStby:=tsSet;
			tModeDuration:=ExDuration_Default_LineStandby;
END_CASE
tModeTime:=TO_TIME(SYSTEMTIME_TO_DT(stSystemTime)-SYSTEMTIME_TO_DT(tsStateChange_local));
m_Set_TimeToExpirationMode:=tModeDuration-tModeTime;

CASE eExTime OF
	E_ExTime.eCIP:;
			tsStateChange:=tsCIP;
	E_ExTime.eWater:;
			tsStateChange:=tsWater;
	E_ExTime.eProduct:;
			tsStateChange:=tsProduction;			
	E_ExTime.eLine :;
			tsStateChange:=tsProductionLine;
	E_ExTime.eLineStby:;
			tsStateChange:=tsProductionLineStby;
END_CASE
END_METHOD

METHOD m_StateUpdate_Limit : BOOL
VAR_INPUT
	value: BOOL;
END_VAR
IF value THEN;
	bStateUpdate_Limited:=TRUE;
ELSE;
	bStateUpdate_Limited:=FALSE;
END_IF
END_METHOD

METHOD m_TimeExpiered : BOOL
VAR_INPUT
END_VAR
CASE eType OF
	E_Element_Type.eTank:;			
	E_Element_Type.eTriBlender:;
	E_Element_Type.eLine:;
	
END_CASE
	
// Rolling Down option
CASE eInterConnect OF
	E_InterConnection.NotConnected:;
				m_TimeExpiredState_RollDown();
	E_InterConnection.ConnToCIP:;
				//do nothing
	E_InterConnection.ConnToLine,
	E_InterConnection.ConnToTriBlender:;
				// Type Tank
				m_TimeExpiredState_RollDown();
	E_InterConnection.ConnToTank:;
				//do nothing
	
END_CASE
END_METHOD

METHOD m_TimeExpiredState_RollDown : BOOL
VAR_INPUT
END_VAR
CASE eState_Long OF
	E_Element_State_Long.eCIP_1_Rinzed:;
				//
	E_Element_State_Long.eCIP_2_Deterged,
	E_Element_State_Long.eCIP_3_Deterged_Clean,
	E_Element_State_Long.eCIP_4_Sanitized,
	E_Element_State_Long.eCIP_5_Done:;	
				State:=E_Element_State_Long.eCIP_1_Rinzed;
	E_Element_State_Long.eWaterReady,
	E_Element_State_Long.eReady,
	E_Element_State_Long.eProduction,
	E_Element_State_Long.eEmpty:;	
			IF eType=E_Element_Type.eTank THEN;
				//State:=E_Element_State_Long.eExpired;
				CASE eElementID OF 
					E_Element_List.eTank_1:;
						IF fbTank1.bReady THEN;
							State:=E_Element_State_Long.eExpired;
						END_IF
						
					E_Element_List.eTank_2:;
						IF fbTank2.bReady THEN;
							State:=E_Element_State_Long.eExpired;
						END_IF
						
					E_Element_List.eTank_3:;
						IF fbTank3.bReady THEN;
							State:=E_Element_State_Long.eExpired;
						END_IF
						
					E_Element_List.eTank_4:;
						IF fbTank4.bReady THEN;
							State:=E_Element_State_Long.eExpired;
						END_IF
												
				END_CASE
				
			ELSE;
				State:=E_Element_State_Long.eNotClean;
			END_IF
			
		E_Element_State_Long.eExpired:;
				IF eType=E_Element_Type.eLine OR eType=E_Element_Type.eTriBlender THEN;
					State:=E_Element_State_Long.eNotClean;
				END_IF
END_CASE
END_METHOD

METHOD m_TimeToExpiration : BOOL
VAR_INPUT
END_VAR
IF tExpirationTime>tStateTime THEN;
	tTimeToExpiration:=tExpirationTime-tStateTime;
ELSE;
	tTimeToExpiration:=T#0S;
	IF TRUE 
	AND eFilling_State=E_Filling_State.eFilling_InProcess
	AND eType=E_Element_Type.eTank
	AND eInterConnect <> E_InterConnection.NotConnected
	AND TRUE
	THEN;
		//Production filling in process 
	ELSE;
		m_TimeExpiered();
	END_IF
	
END_IF

IF State=E_Element_State_Long.eExpired THEN;
	m_TimeExpiered();	
END_IF

IF State=E_Element_State_Long.eStandby 
OR State=E_Element_State_Long.eNotClean
THEN;
	tTimeToExpiration:=T#0S;
END_IF


CASE eType OF
	E_Element_Type.eTank:;		
			CASE eState_Short OF
				E_Element_State_Short.eNotClean:;
						ExpirationTime:=ExDuration_Default;
						eExTime:=E_ExTime.eCIP;
				E_Element_State_Short.eClean:;
						IF eState_Long=E_Element_State_Long.eWaterReady 
						OR (eState_Long=E_Element_State_Long.eExpired
							AND eState_Long_Expiered=E_Element_State_Long.eWaterReady)
						THEN;
							ExpirationTime:=ExDuration_Water;
							eExTime:=E_ExTime.eWater;
						ELSE;
							ExpirationTime:=ExDuration_Default;
							eExTime:=E_ExTime.eCIP;
						END_IF
				E_Element_State_Short.eProduct:;
						ExpirationTime:=ExDuration_Product;
						eExTime:=E_ExTime.eProduct;
			END_CASE			
			
	E_Element_Type.eTriBlender,
	E_Element_Type.eLine:;
			CASE eInterConnect OF
				E_InterConnection.NotConnected:;
					CASE eState_Short OF
						E_Element_State_Short.eNotClean,
						E_Element_State_Short.eClean:;
								ExpirationTime:=ExDuration_Default;
								eExTime:=E_ExTime.eCIP;
	
						E_Element_State_Short.eProduct:;
								IF m_Get_TimeToExpirationMode(eExTime_check:=E_ExTime.eLine)<ExDuration_Default_LineStandby THEN; // line remain time less then 2 hours
									ExpirationTime:=ExDuration_Default_Line;
									eExTime:=E_ExTime.eLine;
								ELSE;
									ExpirationTime:=ExDuration_Default_LineStandby;
									eExTime:=E_ExTime.eLineStby;
								END_IF								
					END_CASE
			
				E_InterConnection.ConnToCIP:;
						ExpirationTime:=ExDuration_Default;
						eExTime:=E_ExTime.eCIP;
						
				E_InterConnection.ConnToTank:;
					CASE eState_Short OF
						E_Element_State_Short.eNotClean,
						E_Element_State_Short.eClean:;
								ExpirationTime:=ExDuration_Default;
								eExTime:=E_ExTime.eCIP;
	
						E_Element_State_Short.eProduct:;		
								ExpirationTime:=ExDuration_Default_Line;
								eExTime:=E_ExTime.eLine;				
					END_CASE
	
						
			ELSE;
		END_CASE
END_CASE


CASE eExTime OF
	E_ExTime.eCIP:;
			tsStateChange:=tsCIP;
	E_ExTime.eWater:;
			tsStateChange:=tsWater;
	E_ExTime.eProduct:;
			tsStateChange:=tsProduction;			
	E_ExTime.eLine :;
			tsStateChange:=tsProductionLine;
	E_ExTime.eLineStby:;
			tsStateChange:=tsProductionLineStby;
END_CASE

CASE eInterConnect OF
	E_InterConnection.NotConnected:;
	E_InterConnection.ConnToCIP:;
	E_InterConnection.ConnToTank:;
	E_InterConnection.ConnToLine:;
	E_InterConnection.ConnToTriBlender:;
END_CASE
END_METHOD

PROPERTY pFilling_State : E_Filling_State
GET
pFilling_State:=eFilling_State;
END_GET
SET
eFilling_State:=pFilling_State;
END_SET
END_PROPERTY

PROPERTY ProdStatus : E_Prod_Status
GET
ProdStatus:=eProdStatus;
END_GET
SET
eProdStatus:=ProdStatus;
END_SET
END_PROPERTY

PROPERTY State : E_Element_State_Long
GET
State:=eState_Long;
END_GET
SET
eState_Long:=State;
END_SET
END_PROPERTY

PROPERTY StateTime : TIMESTRUCT
GET
StateTime:=tsStateChange;
END_GET
SET

CASE eState_Long OF 
	E_Element_State_Long.eOff..			
	E_Element_State_Long.eCIP_5_Done:;
				tsStateChange:=StateTime;
				
				
	//E_Element_State_Long.eOff:;
	//E_Element_State_Long.eOff:;
	//E_Element_State_Long.eOff:;
	
END_CASE
END_SET
END_PROPERTY

END_FUNCTION_BLOCK

// ---- 03 Project/10 Element/FB_Event_echo.TcPOU
FUNCTION_BLOCK FB_Event_echo // for HMI event pudate purpose
VAR_INPUT
END_VAR
VAR_OUTPUT
	echo: INT;
END_VAR
VAR
	ton_time: TON;
	Puls: INT;
	
	memo: BOOL;

END_VAR

ton_time(PT:=T#2S,IN:=memo AND NOT ton_time.Q);
IF ton_time.Q THEN;
	echo:=echo+1;
	
	IF Puls>=5 THEN;
		memo:=FALSE;
	ELSE;
		Puls:=Puls+1;
	END_IF
END_IF

IF ton_time.Q THEN;
	ton_time.IN:=FALSE;
END_IF

METHOD event : BOOL
VAR_INPUT
END_VAR
memo:=TRUE;
echo:=0;
Puls:=0;
END_METHOD

END_FUNCTION_BLOCK

// ---- 03 Project/23 CIP/FB_CIP_Source.TcPOU
FUNCTION_BLOCK FB_CIP_Source EXTENDS FB_SFC_Cycle IMPLEMENTS ITF_FB_SFC_Cycle
VAR_INPUT
	//eElementID			: E_Element_List;
	
	valTank_Water			: E_Pis_Name;
	valTank_R_Water			: E_Pis_Name;
	valTank_Detergent		: E_Pis_Name;
	valTank_DisInfection	: E_Pis_Name;	
	valDrain				: E_Pis_Name;
END_VAR
VAR_OUTPUT
END_VAR
VAR
	//refElement		: REFERENCE TO FB_Element;
	//refState_Long		: REFERENCE TO E_Element_State_Long;
	eReq				: E_CIP_Source;
	eProcess			: E_CIP_Source;
	eStatus				: E_CIP_Source;
	
	fbPis					: FB_Piston;
	stPis_Tank_Water		: REFERENCE TO ST_Piston;
	stPis_Tank_R_Water		: REFERENCE TO ST_Piston;
	stPis_Tank_Detergent	: REFERENCE TO ST_Piston;
	stPis_Tank_DisInfection	: REFERENCE TO ST_Piston;
	stPis_Drain				: REFERENCE TO ST_Piston;
	rt_Req_Reset: R_TRIG;
END_VAR
VAR_IN_OUT


END_VAR

act_GetReference();

act_Oper();
IF NOT Init.x THEN;
	act_Status();
END_IF

m_Request_Reset(memo:=rt_Req_Reset);//

ACTION _aClose_active:
bStepDone:=FALSE;
IF TRUE 
AND eStatus=E_CIP_Source.eClose
THEN;
	bStepDone:=TRUE;
END_IF
END_ACTION

ACTION _aClose_entry:
fbPis.m_SetByRecipe(stPis:=stPis_Tank_Water, 			req:=E_Piston_Recipe_State.Release);
fbPis.m_SetByRecipe(stPis:=stPis_Tank_R_Water, 			req:=E_Piston_Recipe_State.Release);
fbPis.m_SetByRecipe(stPis:=stPis_Tank_Detergent, 		req:=E_Piston_Recipe_State.Release);
fbPis.m_SetByRecipe(stPis:=stPis_Tank_DisInfection, 	req:=E_Piston_Recipe_State.Release);
fbPis.m_SetByRecipe(stPis:=stPis_Drain, 				req:=E_Piston_Recipe_State.Release);
END_ACTION

ACTION _aDetergent_entry:
fbPis.m_SetByRecipe(stPis:=stPis_Tank_Water, 			req:=E_Piston_Recipe_State.Release);
fbPis.m_SetByRecipe(stPis:=stPis_Tank_R_Water, 			req:=E_Piston_Recipe_State.Release);
fbPis.m_SetByRecipe(stPis:=stPis_Tank_Detergent, 		req:=E_Piston_Recipe_State.Act);
fbPis.m_SetByRecipe(stPis:=stPis_Tank_DisInfection, 	req:=E_Piston_Recipe_State.Release);
//fbPis.m_SetByRecipe(stPis:=stPis_Drain, 				req:=E_Piston_Recipe_State.Act);
END_ACTION

ACTION _aDone_entry:
eProcess:=E_CIP_Source.eNone;
eReq:=E_CIP_Source.eNone;
bRun:=FALSE;
bDone:=TRUE;
END_ACTION

ACTION _aInit_active:
SFCReset:=FALSE;
END_ACTION

ACTION _aInit_exit:
eProcess:=E_CIP_Source.eNone;
eReq:=E_CIP_Source.eNone;
END_ACTION

ACTION _aR_Water_entry:
fbPis.m_SetByRecipe(stPis:=stPis_Tank_Water, 			req:=E_Piston_Recipe_State.Release);
fbPis.m_SetByRecipe(stPis:=stPis_Tank_R_Water, 			req:=E_Piston_Recipe_State.Act);
fbPis.m_SetByRecipe(stPis:=stPis_Tank_Detergent, 		req:=E_Piston_Recipe_State.Release);
fbPis.m_SetByRecipe(stPis:=stPis_Tank_DisInfection, 	req:=E_Piston_Recipe_State.Release);
//fbPis.m_SetByRecipe(stPis:=stPis_Drain, 				req:=E_Piston_Recipe_State.Act);
END_ACTION

ACTION _aReady_active:


CASE eReq OF
	E_CIP_Source.eClose:;
			IF TRUE THEN;
				eProcess:=E_CIP_Source.eClose;
			END_IF

	E_CIP_Source.eT91_Sanitation:;
			IF TRUE THEN;
				eProcess:=E_CIP_Source.eT91_Sanitation;
			END_IF	
			
	E_CIP_Source.eT92_Detergent:;
			IF TRUE THEN;
				eProcess:=E_CIP_Source.eT92_Detergent;
			END_IF	

	E_CIP_Source.eT93_R_Water:;
			IF TRUE THEN;
				eProcess:=E_CIP_Source.eT93_R_Water;
			END_IF	
			
	E_CIP_Source.eT94_Water:;
			IF TRUE THEN;
				eProcess:=E_CIP_Source.eT94_Water;
			END_IF	

END_CASE
END_ACTION

ACTION _aReady_entry:

END_ACTION

ACTION _aReady_exit:
bRun:=TRUE;
bDone:=FALSE;
END_ACTION

ACTION _aSanitation_entry:
fbPis.m_SetByRecipe(stPis:=stPis_Tank_Water, 			req:=E_Piston_Recipe_State.Release);
fbPis.m_SetByRecipe(stPis:=stPis_Tank_R_Water, 			req:=E_Piston_Recipe_State.Release);
fbPis.m_SetByRecipe(stPis:=stPis_Tank_Detergent, 		req:=E_Piston_Recipe_State.Release);
fbPis.m_SetByRecipe(stPis:=stPis_Tank_DisInfection, 	req:=E_Piston_Recipe_State.Act);
END_ACTION

ACTION _aT91_Drain_Done_active:
bStepDone:=FALSE;
IF TRUE 
AND eStatus=E_CIP_Source.eT91_Sanitation
THEN;
	bStepDone:=TRUE;
END_IF
END_ACTION

ACTION _aT91_Drain_Done_entry:
fbPis.m_SetByRecipe(stPis:=stPis_Drain, 				req:=E_Piston_Recipe_State.Act);
END_ACTION

ACTION _aT92_Drain_Done_active:
bStepDone:=FALSE;
IF TRUE 
AND eStatus=E_CIP_Source.eT92_Detergent
THEN;
	bStepDone:=TRUE;
END_IF
END_ACTION

ACTION _aT92_Drain_Done_entry:
fbPis.m_SetByRecipe(stPis:=stPis_Drain, 				req:=E_Piston_Recipe_State.Act);
END_ACTION

ACTION _aT93_Drain_Done_active:
bStepDone:=FALSE;
IF TRUE 
AND eStatus=E_CIP_Source.eT93_R_Water
THEN;
	bStepDone:=TRUE;
END_IF
END_ACTION

ACTION _aT93_Drain_Done_entry:
fbPis.m_SetByRecipe(stPis:=stPis_Drain, 				req:=E_Piston_Recipe_State.Act);
END_ACTION

ACTION _aWater_active:
bStepDone:=FALSE;
IF TRUE 
AND eStatus=E_CIP_Source.eT94_Water
THEN;
	bStepDone:=TRUE;
END_IF
END_ACTION

ACTION _aWater_entry:
fbPis.m_SetByRecipe(stPis:=stPis_Tank_Water, 			req:=E_Piston_Recipe_State.Act);
fbPis.m_SetByRecipe(stPis:=stPis_Tank_R_Water, 			req:=E_Piston_Recipe_State.Release);
fbPis.m_SetByRecipe(stPis:=stPis_Tank_Detergent, 		req:=E_Piston_Recipe_State.Release);
fbPis.m_SetByRecipe(stPis:=stPis_Tank_DisInfection, 	req:=E_Piston_Recipe_State.Release);
fbPis.m_SetByRecipe(stPis:=stPis_Drain, 				req:=E_Piston_Recipe_State.Release);
END_ACTION

ACTION act_GetReference:
m_Set_SFCFlags_Reference();
//refElement REF= fbElement[eElementID];
//refState_Long REF= fbElement[eElementID].eState_Long;
	
stPis_Tank_Water			REF= g_Piston.stPis[valTank_Water];
stPis_Tank_R_Water			REF= g_Piston.stPis[valTank_R_Water];
stPis_Tank_Detergent		REF= g_Piston.stPis[valTank_Detergent];
stPis_Tank_DisInfection		REF= g_Piston.stPis[valTank_DisInfection];
stPis_Drain					REF= g_Piston.stPis[valDrain];
END_ACTION

ACTION act_Oper:
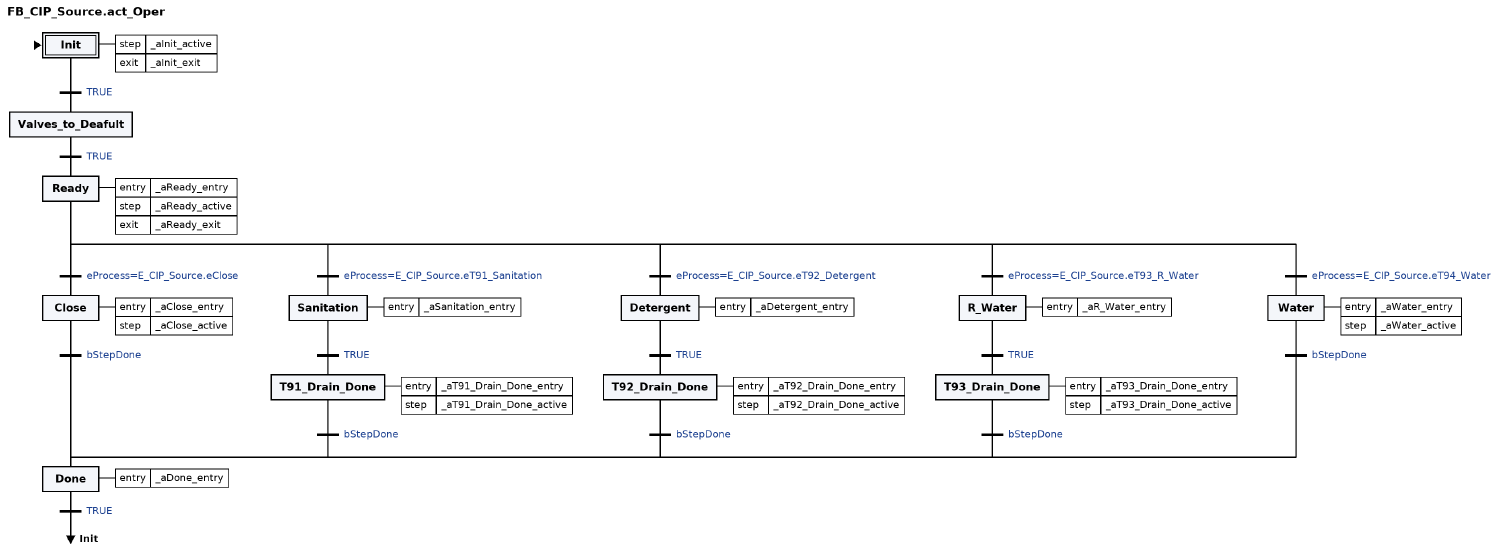
INITIAL_STEP Init:  // min time T#0.5s
    _aInit_active(N);  // step action
    _aInit_exit(P0);  // exit action
END_STEP
TRANSITION FROM Init TO Valves_to_Deafult
    := TRUE;
END_TRANSITION
STEP Valves_to_Deafult:
END_STEP
TRANSITION FROM Valves_to_Deafult TO Ready
    := TRUE;
END_TRANSITION
STEP Ready:
    _aReady_entry(P1);  // entry action
    _aReady_active(N);  // step action
    _aReady_exit(P0);  // exit action
END_STEP
TRANSITION FROM Ready TO Close
    := eProcess=E_CIP_Source.eClose;
END_TRANSITION
STEP Close:
    _aClose_entry(P1);  // entry action
    _aClose_active(N);  // step action
END_STEP
TRANSITION FROM Close TO Done
    := bStepDone;
END_TRANSITION
TRANSITION FROM Ready TO Sanitation
    := eProcess=E_CIP_Source.eT91_Sanitation;
END_TRANSITION
STEP Sanitation:  // min time T#7s
    _aSanitation_entry(P1);  // entry action
END_STEP
TRANSITION FROM Sanitation TO T91_Drain_Done
    := TRUE;
END_TRANSITION
STEP T91_Drain_Done:
    _aT91_Drain_Done_entry(P1);  // entry action
    _aT91_Drain_Done_active(N);  // step action
END_STEP
TRANSITION FROM T91_Drain_Done TO Done
    := bStepDone;
END_TRANSITION
TRANSITION FROM Ready TO Detergent
    := eProcess=E_CIP_Source.eT92_Detergent;
END_TRANSITION
STEP Detergent:  // min time T#6s
    _aDetergent_entry(P1);  // entry action
END_STEP
TRANSITION FROM Detergent TO T92_Drain_Done
    := TRUE;
END_TRANSITION
STEP T92_Drain_Done:
    _aT92_Drain_Done_entry(P1);  // entry action
    _aT92_Drain_Done_active(N);  // step action
END_STEP
TRANSITION FROM T92_Drain_Done TO Done
    := bStepDone;
END_TRANSITION
TRANSITION FROM Ready TO R_Water
    := eProcess=E_CIP_Source.eT93_R_Water;
END_TRANSITION
STEP R_Water:  // min time T#5s
    _aR_Water_entry(P1);  // entry action
END_STEP
TRANSITION FROM R_Water TO T93_Drain_Done
    := TRUE;
END_TRANSITION
STEP T93_Drain_Done:
    _aT93_Drain_Done_entry(P1);  // entry action
    _aT93_Drain_Done_active(N);  // step action
END_STEP
TRANSITION FROM T93_Drain_Done TO Done
    := bStepDone;
END_TRANSITION
TRANSITION FROM Ready TO Water
    := eProcess=E_CIP_Source.eT94_Water;
END_TRANSITION
STEP Water:
    _aWater_entry(P1);  // entry action
    _aWater_active(N);  // step action
END_STEP
TRANSITION FROM Water TO Done
    := bStepDone;
END_TRANSITION
STEP Done:  // min time T#0.2s
    _aDone_entry(P1);  // entry action
END_STEP
TRANSITION FROM Done TO Init
    := TRUE;
END_TRANSITION
// branch label Branch1_act_Oper
END_ACTION

ACTION act_Status:
IF bReady AND bDone OR TRUE THEN;
	IF TRUE 
	AND fbPis.m_CheckByRecipe(stPis:=stPis_Tank_Water, 			req:=E_Piston_Recipe_State.Release)
	AND fbPis.m_CheckByRecipe(stPis:=stPis_Tank_R_Water, 		req:=E_Piston_Recipe_State.Release)
	AND fbPis.m_CheckByRecipe(stPis:=stPis_Tank_Detergent, 		req:=E_Piston_Recipe_State.Release)
	AND fbPis.m_CheckByRecipe(stPis:=stPis_Tank_DisInfection, 	req:=E_Piston_Recipe_State.Release)
	AND fbPis.m_CheckByRecipe(stPis:=stPis_Drain, 				req:=E_Piston_Recipe_State.Release)
	THEN;
		eStatus:=E_CIP_Source.eClose;
	
	ELSIF TRUE 
	AND fbPis.m_CheckByRecipe(stPis:=stPis_Tank_Water, 			req:=E_Piston_Recipe_State.Act)
	AND fbPis.m_CheckByRecipe(stPis:=stPis_Tank_R_Water, 		req:=E_Piston_Recipe_State.Release)
	AND fbPis.m_CheckByRecipe(stPis:=stPis_Tank_Detergent, 		req:=E_Piston_Recipe_State.Release)
	AND fbPis.m_CheckByRecipe(stPis:=stPis_Tank_DisInfection, 	req:=E_Piston_Recipe_State.Release)
	AND fbPis.m_CheckByRecipe(stPis:=stPis_Drain, 				req:=E_Piston_Recipe_State.Release)
	THEN;
		eStatus:=E_CIP_Source.eT94_Water;
		
	ELSIF TRUE 
	AND fbPis.m_CheckByRecipe(stPis:=stPis_Tank_Water, 			req:=E_Piston_Recipe_State.Release)
	AND fbPis.m_CheckByRecipe(stPis:=stPis_Tank_R_Water, 		req:=E_Piston_Recipe_State.Act)
	AND fbPis.m_CheckByRecipe(stPis:=stPis_Tank_Detergent, 		req:=E_Piston_Recipe_State.Release)
	AND fbPis.m_CheckByRecipe(stPis:=stPis_Tank_DisInfection, 	req:=E_Piston_Recipe_State.Release)
	AND fbPis.m_CheckByRecipe(stPis:=stPis_Drain, 				req:=E_Piston_Recipe_State.Act)
	THEN;
		eStatus:=E_CIP_Source.eT93_R_Water;
		
	ELSIF TRUE 	
	AND fbPis.m_CheckByRecipe(stPis:=stPis_Tank_Water, 			req:=E_Piston_Recipe_State.Release)
	AND fbPis.m_CheckByRecipe(stPis:=stPis_Tank_R_Water, 		req:=E_Piston_Recipe_State.Release)
	AND fbPis.m_CheckByRecipe(stPis:=stPis_Tank_Detergent, 		req:=E_Piston_Recipe_State.Act)
	AND fbPis.m_CheckByRecipe(stPis:=stPis_Tank_DisInfection, 	req:=E_Piston_Recipe_State.Release)
	AND fbPis.m_CheckByRecipe(stPis:=stPis_Drain, 				req:=E_Piston_Recipe_State.Act)
	THEN;
		eStatus:=E_CIP_Source.eT92_Detergent;
		
	ELSIF TRUE 	
	AND fbPis.m_CheckByRecipe(stPis:=stPis_Tank_Water, 			req:=E_Piston_Recipe_State.Release)
	AND fbPis.m_CheckByRecipe(stPis:=stPis_Tank_R_Water, 		req:=E_Piston_Recipe_State.Release)
	AND fbPis.m_CheckByRecipe(stPis:=stPis_Tank_Detergent, 		req:=E_Piston_Recipe_State.Release)
	AND fbPis.m_CheckByRecipe(stPis:=stPis_Tank_DisInfection, 	req:=E_Piston_Recipe_State.Act)
	AND fbPis.m_CheckByRecipe(stPis:=stPis_Drain, 				req:=E_Piston_Recipe_State.Act)
	THEN;
		eStatus:=E_CIP_Source.eT91_Sanitation;
	ELSE;
		eStatus:=E_Tank_Target.eNone;
	END_IF
ELSE;
	eStatus:=E_Tank_Target.eNone;
END_IF
END_ACTION

METHOD m_CheckStatus : BOOL
VAR_INPUT
	eReqStatus		: E_CIP_Source;
END_VAR
IF eStatus=eReqStatus 
AND eProcess=E_CIP_Source.eNone
AND eReq=E_CIP_Source.eNone
AND bReady
AND bDone
AND NOT bRun
THEN;
	m_CheckStatus:=TRUE;
END_IF
END_METHOD

METHOD m_Request_Reset : BOOL
VAR_IN_OUT
	memo: R_TRIG;
END_VAR
memo(CLK:=eReq=0);
IF TRUE 
AND memo.Q
THEN;
	SFCReset:=TRUE;
END_IF
END_METHOD

METHOD m_Run : BOOL
VAR_INPUT
	eReqProc			: E_CIP_Source;
END_VAR
IF eProcess=E_CIP_Source.eNone THEN;
	eProcess:=eReq:=eReqProc;
	bDone:=FALSE;
	m_Run:=TRUE;
END_IF
END_METHOD

METHOD m_Set_SFCFlags_Reference : BOOL
//Set reference to SFC flags

refSFC.SFCInit REF= SFCInit;
refSFC.SFCReset REF= SFCReset;
refSFC.SFCError REF= SFCError;
refSFC.SFCEnableLimit REF= SFCEnableLimit;
refSFC.SFCErrorStep REF= SFCErrorStep;
refSFC.SFCErrorPOU REF= SFCErrorPOU;
refSFC.SFCQuitError REF= SFCQuitError;
refSFC.SFCPause REF= SFCPause;
refSFC.SFCTrans REF= SFCTrans;
refSFC.SFCCurrentStep REF= SFCCurrentStep;
refSFC.SFCTip REF= SFCTip;
refSFC.SFCTipMode REF= SFCTipMode;

// Cycle handle for SFC
m_SFC_Handle();
END_METHOD

END_FUNCTION_BLOCK

// ---- 00 Library/03 SFC/FB_SFC_Cycle.TcPOU
FUNCTION_BLOCK FB_SFC_Cycle
VAR_INPUT

END_VAR
VAR_OUTPUT
END_VAR
VAR
	refSFC: ST_SFC;

	bInit: BOOL;
	bResetCycle: BOOL;
	bResume: BOOL;
	bRun: BOOL;	
	bReady: BOOL;
	bDone: BOOL;
	bToBe_Done: BOOL;
	
	bStepMode: BOOL;
	bNextStep: BOOL;



	bStepDone: BOOL;
	ton_StepTime: TON;
	
	StageDelayByRecipe: TIME;
	
	//fbPis_Meth: FB_Piston;

	rtDone	: R_TRIG;
	rtRun	: R_TRIG;
	sLastStepBefore_Error	: STRING;
	sError_Message			: STRING;
	
	ErrorSFC: BOOL;

	tonResetCycle: TON;
	
	stMode_zone	: REFERENCE TO ST_Mode;
	stOper_zone	: REFERENCE TO ST_OperationButtons;
	ftStateSafe : F_TRIG;
	
END_VAR

METHOD m_Reset_LastStepBeforeError : BOOL
VAR_INPUT
END_VAR
sLastStepBefore_Error:='';
END_METHOD

METHOD m_Set_LastStepBeforeError : BOOL
VAR_INPUT
END_VAR
sLastStepBefore_Error:=refSFC.SFCCurrentStep;
END_METHOD

METHOD m_Set_Mode_Reference : BOOL
VAR_INPUT
	inMoedeZone: E_ModeZone;
END_VAR
stMode_zone REF=(stMode[inMoedeZone]);
stOper_zone REF=(stOper[inMoedeZone]);
END_METHOD

METHOD m_SFC_Handle : BOOL
VAR_INPUT
END_VAR

VAR
	
END_VAR
IF NOT __ISVALIDREF(refSFC.SFCInit) 
OR NOT  __ISVALIDREF(refSFC.SFCReset) 
OR NOT  __ISVALIDREF(refSFC.SFCError) 
OR NOT  __ISVALIDREF(refSFC.SFCEnableLimit) 
OR NOT  __ISVALIDREF(refSFC.SFCErrorStep) 
OR NOT  __ISVALIDREF(refSFC.SFCErrorPOU) 
OR NOT  __ISVALIDREF(refSFC.SFCQuitError) 
OR NOT  __ISVALIDREF(refSFC.SFCPause) 
OR NOT  __ISVALIDREF(refSFC.SFCTrans) 
OR NOT  __ISVALIDREF(refSFC.SFCCurrentStep) 
OR NOT  __ISVALIDREF(refSFC.SFCTip) 
OR NOT  __ISVALIDREF(refSFC.SFCTipMode) 
THEN;
	RETURN;
END_IF

refSFC.SFCEnableLimit:=TRUE;
IF refSFC.SFCTrans THEN;
	bStepDone:=FALSE;
	ton_StepTime(IN:=FALSE);
ELSE;
	ton_StepTime(IN:=TRUE); //depend on step condition
END_IF

IF bInit THEN;
	refSFC.SFCInit:=TRUE;
ELSE;
	refSFC.SFCInit:=FALSE;
END_IF

IF refSFC.SFCError THEN;
	refSFC.SFCPause:=TRUE;
	ErrorSFC:=TRUE;
	m_Set_LastStepBeforeError();
END_IF

IF refSFC.SFCQuitError THEN;
	refSFC.SFCPause:=FALSE;
	ErrorSFC:=FALSE;
	refSFC.SFCQuitError:=FALSE;
	m_Reset_LastStepBeforeError();
	sError_Message:='';
END_IF

IF refSFC.SFCCurrentStep='Ready' THEN;
	bReady:=TRUE;
ELSE;
	bReady:=FALSE;
END_IF

rtDone(CLK:=refSFC.SFCCurrentStep='Done');
IF rtDone.Q THEN;
	bDone:=TRUE;
END_IF
rtRun(CLK:=bRun);
IF rtRun.Q THEN;
	bDone:=FALSE;
END_IF

IF bResume THEN;
	ErrorSFC:=FALSE;
	refSFC.SFCError:=FALSE;
	refSFC.SFCPause:=FALSE;
	m_Reset_LastStepBeforeError();
	bResume:=FALSE;
END_IF


tonResetCycle(PT:=T#0.5S,IN:=bResetCycle);
IF bResetCycle THEN;
	refSFC.SFCReset:=TRUE;
	//tonResetCycle.IN:=TRUE;
END_IF
IF tonResetCycle.Q THEN;
	bResetCycle:=FALSE;
	refSFC.SFCReset:=FALSE;
END_IF

StepByStep();

IF NOT __ISVALIDREF(stMode_zone)
OR NOT __ISVALIDREF(stOper_zone)
THEN;
	RETURN;
ELSE;
	//IF prg_Safety.ftStateSafe.Q THEN;
	ftStateSafe(CLK:=stMode_zone.bStateSafe_mode);
	IF ftStateSafe.Q THEN;
		//bResetCycle:=TRUE;
	END_IF	
END_IF



(*
rtDone(CLK:=bDone);
IF rtDone.Q THEN
	bToBe_Done:=FALSE;
END_IF
*)
END_METHOD

METHOD mInit : BOOL
VAR_INPUT
END_VAR
bInit:=TRUE;
bToBe_Done:=FALSE;
END_METHOD

METHOD mResetCycle : BOOL
VAR_INPUT
END_VAR
bResetCycle:=TRUE;
bRun:=FALSE;
refSFC.SFCReset:=TRUE;
END_METHOD

METHOD mRun : BOOL
VAR_INPUT
	
END_VAR
bRun:=TRUE;
bDone:=FALSE;

IF rtDone.Q THEN;
	mRun:=TRUE;	
END_IF
END_METHOD

METHOD mToBe_Done : BOOL
VAR_INPUT
END_VAR
bToBe_Done:=TRUE;
bDone:=FALSE;
END_METHOD

METHOD StepByStep : BOOL
VAR_INPUT
END_VAR


IF bStepMode THEN;
	IF refSFC.SFCTrans THEN;
		refSFC.SFCTipMode:=TRUE;
		bNextStep:=FALSE;
	END_IF
	IF bNextStep THEN;
		refSFC.SFCTipMode:=FALSE;
	END_IF
ELSE;
	refSFC.SFCTipMode:=FALSE;
END_IF
END_METHOD

END_FUNCTION_BLOCK

// ---- 03 Project/23 CIP/FB_CIP_Return.TcPOU
FUNCTION_BLOCK FB_CIP_Return EXTENDS FB_SFC_Cycle IMPLEMENTS ITF_FB_SFC_Cycle
VAR_INPUT
	//eElementID			: E_Element_List;
	
	valTank_Water			: E_Pis_Name;
	valTank_Water_1			: E_Pis_Name;
	valTank_R_Water			: E_Pis_Name;
	valTank_R_Water_1		: E_Pis_Name;
	valTank_Detergent		: E_Pis_Name;
	valTank_Detergent_1		: E_Pis_Name;
	valTank_DisInfection	: E_Pis_Name;
	valTank_DisInfection_1	: E_Pis_Name;
	valDrain				: E_Pis_Name;
	
END_VAR
VAR_OUTPUT
END_VAR
VAR
	//refElement		: REFERENCE TO FB_Element;
	//refState_Long		: REFERENCE TO E_Element_State_Long;
	eReq				: E_CIP_Return;
	eProcess			: E_CIP_Return;
	eStatus				: E_CIP_Return;
	
	fbPis						: FB_Piston;
	stPis_Tank_Water			: REFERENCE TO ST_Piston;
	stPis_Tank_Water_1			: REFERENCE TO ST_Piston;
	stPis_Tank_R_Water			: REFERENCE TO ST_Piston;
	stPis_Tank_R_Water_1		: REFERENCE TO ST_Piston;
	stPis_Tank_Detergent		: REFERENCE TO ST_Piston;
	stPis_Tank_Detergent_1		: REFERENCE TO ST_Piston;
	stPis_Tank_DisInfection		: REFERENCE TO ST_Piston;
	stPis_Tank_DisInfection_1	: REFERENCE TO ST_Piston;
	stPis_Drain					: REFERENCE TO ST_Piston;
	rt_Req_Reset: R_TRIG;
END_VAR
VAR_IN_OUT


END_VAR

act_GetReference();

act_Oper();
IF NOT Init.x THEN;
	act_Status();
END_IF

m_Request_Reset(memo:=rt_Req_Reset);//

ACTION _aDetergent_active:
bStepDone:=FALSE;
IF TRUE 
AND eStatus=E_CIP_Return.eT92_Detergent
THEN;
	bStepDone:=TRUE;
END_IF
END_ACTION

ACTION _aDetergent_entry:
fbPis.m_SetByRecipe(stPis:=stPis_Tank_Water, 			req:=E_Piston_Recipe_State.Release);
fbPis.m_SetByRecipe(stPis:=stPis_Tank_Water_1, 			req:=E_Piston_Recipe_State.Release);
fbPis.m_SetByRecipe(stPis:=stPis_Tank_R_Water, 			req:=E_Piston_Recipe_State.Release);
fbPis.m_SetByRecipe(stPis:=stPis_Tank_R_Water_1, 		req:=E_Piston_Recipe_State.Release);
fbPis.m_SetByRecipe(stPis:=stPis_Tank_Detergent, 		req:=E_Piston_Recipe_State.Act);
fbPis.m_SetByRecipe(stPis:=stPis_Tank_Detergent_1, 		req:=E_Piston_Recipe_State.Act);
fbPis.m_SetByRecipe(stPis:=stPis_Tank_DisInfection_1, 	req:=E_Piston_Recipe_State.Release);
fbPis.m_SetByRecipe(stPis:=stPis_Tank_DisInfection, 	req:=E_Piston_Recipe_State.Release);
fbPis.m_SetByRecipe(stPis:=stPis_Drain, 				req:=E_Piston_Recipe_State.Release);
END_ACTION

ACTION _aDone_entry:
eProcess:=E_CIP_Return.eNone; 
eReq:=E_CIP_Return.eNone;
bRun:=FALSE;
bDone:=TRUE;
END_ACTION

ACTION _aDrain_active:
bStepDone:=FALSE;
IF TRUE 
AND eStatus=E_CIP_Return.eDrain
THEN;
	bStepDone:=TRUE;
END_IF
END_ACTION

ACTION _aDrain_entry:
fbPis.m_SetByRecipe(stPis:=stPis_Tank_Water, 			req:=E_Piston_Recipe_State.Release);
fbPis.m_SetByRecipe(stPis:=stPis_Tank_Water_1, 			req:=E_Piston_Recipe_State.Release);
fbPis.m_SetByRecipe(stPis:=stPis_Tank_R_Water, 			req:=E_Piston_Recipe_State.Release);
fbPis.m_SetByRecipe(stPis:=stPis_Tank_R_Water_1, 		req:=E_Piston_Recipe_State.Release);
fbPis.m_SetByRecipe(stPis:=stPis_Tank_Detergent, 		req:=E_Piston_Recipe_State.Release);
fbPis.m_SetByRecipe(stPis:=stPis_Tank_Detergent_1, 		req:=E_Piston_Recipe_State.Release);
fbPis.m_SetByRecipe(stPis:=stPis_Tank_DisInfection, 	req:=E_Piston_Recipe_State.Release);
fbPis.m_SetByRecipe(stPis:=stPis_Tank_DisInfection_1, 	req:=E_Piston_Recipe_State.Release);
fbPis.m_SetByRecipe(stPis:=stPis_Drain, 				req:=E_Piston_Recipe_State.Release);
END_ACTION

ACTION _aInit_active:
SFCReset:=FALSE;
END_ACTION

ACTION _aInit_exit:
eProcess:=E_CIP_Return.eNone;
eReq:=E_CIP_Return.eNone;
END_ACTION

ACTION _aR_Water_active:
bStepDone:=FALSE;
IF TRUE 
AND eStatus=E_CIP_Return.eT93_R_Water
THEN;
	bStepDone:=TRUE;
END_IF
END_ACTION

ACTION _aR_Water_entry:
fbPis.m_SetByRecipe(stPis:=stPis_Tank_Water, 			req:=E_Piston_Recipe_State.Release);
fbPis.m_SetByRecipe(stPis:=stPis_Tank_Water_1, 			req:=E_Piston_Recipe_State.Release);
fbPis.m_SetByRecipe(stPis:=stPis_Tank_R_Water, 			req:=E_Piston_Recipe_State.Act);
fbPis.m_SetByRecipe(stPis:=stPis_Tank_R_Water_1, 		req:=E_Piston_Recipe_State.Act);
fbPis.m_SetByRecipe(stPis:=stPis_Tank_Detergent, 		req:=E_Piston_Recipe_State.Release);
fbPis.m_SetByRecipe(stPis:=stPis_Tank_Detergent_1, 		req:=E_Piston_Recipe_State.Release);
fbPis.m_SetByRecipe(stPis:=stPis_Tank_DisInfection, 	req:=E_Piston_Recipe_State.Release);
fbPis.m_SetByRecipe(stPis:=stPis_Tank_DisInfection_1, 	req:=E_Piston_Recipe_State.Release);
fbPis.m_SetByRecipe(stPis:=stPis_Drain, 				req:=E_Piston_Recipe_State.Release);
END_ACTION

ACTION _aReady_active:


CASE eReq OF
	E_CIP_Return.eDrain:;
			IF TRUE THEN;
				eProcess:=E_CIP_Return.eDrain;
			END_IF

	E_CIP_Return.eT91_Sanitation:;
			IF TRUE THEN;
				eProcess:=E_CIP_Return.eT91_Sanitation;
			END_IF	
			
	E_CIP_Return.eT92_Detergent:;
			IF TRUE THEN;
				eProcess:=E_CIP_Return.eT92_Detergent;
			END_IF	

	E_CIP_Return.eT93_R_Water:;
			IF TRUE THEN;
				eProcess:=E_CIP_Return.eT93_R_Water;
			END_IF	
			
	E_CIP_Return.eT94_Water:;
			IF TRUE THEN;
				eProcess:=E_CIP_Return.eT94_Water;
			END_IF	

END_CASE
END_ACTION

ACTION _aReady_entry:

END_ACTION

ACTION _aReady_exit:
bRun:=TRUE;
bDone:=FALSE;
END_ACTION

ACTION _aSanitation_active:
bStepDone:=FALSE;
IF TRUE 
AND eStatus=E_CIP_Return.eT91_Sanitation
THEN;
	bStepDone:=TRUE;
END_IF
END_ACTION

ACTION _aSanitation_entry:
fbPis.m_SetByRecipe(stPis:=stPis_Tank_Water, 			req:=E_Piston_Recipe_State.Release);
fbPis.m_SetByRecipe(stPis:=stPis_Tank_Water_1, 			req:=E_Piston_Recipe_State.Release);
fbPis.m_SetByRecipe(stPis:=stPis_Tank_R_Water, 			req:=E_Piston_Recipe_State.Release);
fbPis.m_SetByRecipe(stPis:=stPis_Tank_R_Water_1, 		req:=E_Piston_Recipe_State.Release);
fbPis.m_SetByRecipe(stPis:=stPis_Tank_Detergent, 		req:=E_Piston_Recipe_State.Release);
fbPis.m_SetByRecipe(stPis:=stPis_Tank_Detergent_1, 		req:=E_Piston_Recipe_State.Release);
fbPis.m_SetByRecipe(stPis:=stPis_Tank_DisInfection, 	req:=E_Piston_Recipe_State.Act);
fbPis.m_SetByRecipe(stPis:=stPis_Tank_DisInfection_1, 	req:=E_Piston_Recipe_State.Act);
fbPis.m_SetByRecipe(stPis:=stPis_Drain, 				req:=E_Piston_Recipe_State.Release);
END_ACTION

ACTION _aWater_active:
bStepDone:=FALSE;
IF TRUE 
AND eStatus=E_CIP_Return.eT94_Water
THEN;
	bStepDone:=TRUE;
END_IF
END_ACTION

ACTION _aWater_entry:
fbPis.m_SetByRecipe(stPis:=stPis_Tank_Water, 			req:=E_Piston_Recipe_State.Act);
fbPis.m_SetByRecipe(stPis:=stPis_Tank_Water_1, 			req:=E_Piston_Recipe_State.Act);
fbPis.m_SetByRecipe(stPis:=stPis_Tank_R_Water, 			req:=E_Piston_Recipe_State.Release);
fbPis.m_SetByRecipe(stPis:=stPis_Tank_R_Water_1, 		req:=E_Piston_Recipe_State.Release);
fbPis.m_SetByRecipe(stPis:=stPis_Tank_Detergent, 		req:=E_Piston_Recipe_State.Release);
fbPis.m_SetByRecipe(stPis:=stPis_Tank_Detergent_1, 		req:=E_Piston_Recipe_State.Release);
fbPis.m_SetByRecipe(stPis:=stPis_Tank_DisInfection, 	req:=E_Piston_Recipe_State.Release);
fbPis.m_SetByRecipe(stPis:=stPis_Tank_DisInfection_1, 	req:=E_Piston_Recipe_State.Release);
fbPis.m_SetByRecipe(stPis:=stPis_Drain, 				req:=E_Piston_Recipe_State.Act);
END_ACTION

ACTION act_GetReference:
m_Set_SFCFlags_Reference();
//refElement REF= fbElement[eElementID];
//refState_Long REF= fbElement[eElementID].eState_Long;
	
stPis_Tank_Water				REF= g_Piston.stPis[valTank_Water];
stPis_Tank_Water_1				REF= g_Piston.stPis[valTank_Water_1];
stPis_Tank_R_Water				REF= g_Piston.stPis[valTank_R_Water];
stPis_Tank_R_Water_1			REF= g_Piston.stPis[valTank_R_Water_1];
stPis_Tank_Detergent			REF= g_Piston.stPis[valTank_Detergent];
stPis_Tank_Detergent_1			REF= g_Piston.stPis[valTank_Detergent_1];
stPis_Tank_DisInfection			REF= g_Piston.stPis[valTank_DisInfection];
stPis_Tank_DisInfection_1		REF= g_Piston.stPis[valTank_DisInfection_1];
stPis_Drain						REF= g_Piston.stPis[valDrain];
END_ACTION

ACTION act_Oper:
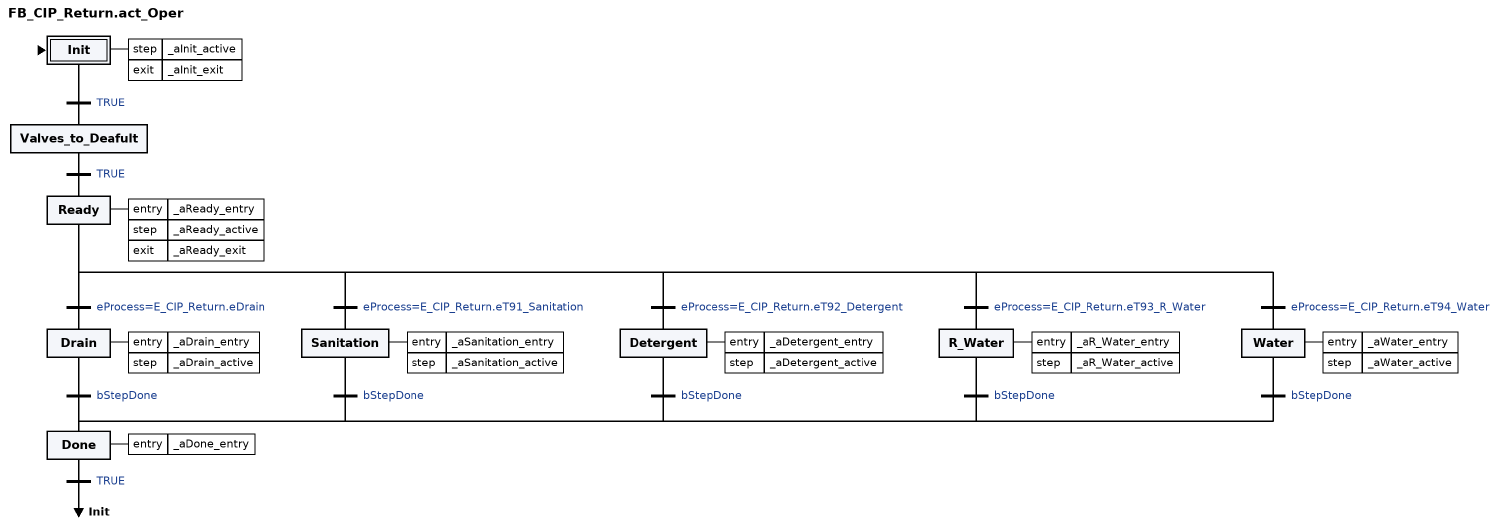
INITIAL_STEP Init:  // min time T#0.5s
    _aInit_active(N);  // step action
    _aInit_exit(P0);  // exit action
END_STEP
TRANSITION FROM Init TO Valves_to_Deafult
    := TRUE;
END_TRANSITION
STEP Valves_to_Deafult:
END_STEP
TRANSITION FROM Valves_to_Deafult TO Ready
    := TRUE;
END_TRANSITION
STEP Ready:
    _aReady_entry(P1);  // entry action
    _aReady_active(N);  // step action
    _aReady_exit(P0);  // exit action
END_STEP
TRANSITION FROM Ready TO Drain
    := eProcess=E_CIP_Return.eDrain;
END_TRANSITION
STEP Drain:
    _aDrain_entry(P1);  // entry action
    _aDrain_active(N);  // step action
END_STEP
TRANSITION FROM Drain TO Done
    := bStepDone;
END_TRANSITION
TRANSITION FROM Ready TO Sanitation
    := eProcess=E_CIP_Return.eT91_Sanitation;
END_TRANSITION
STEP Sanitation:
    _aSanitation_entry(P1);  // entry action
    _aSanitation_active(N);  // step action
END_STEP
TRANSITION FROM Sanitation TO Done
    := bStepDone;
END_TRANSITION
TRANSITION FROM Ready TO Detergent
    := eProcess=E_CIP_Return.eT92_Detergent;
END_TRANSITION
STEP Detergent:
    _aDetergent_entry(P1);  // entry action
    _aDetergent_active(N);  // step action
END_STEP
TRANSITION FROM Detergent TO Done
    := bStepDone;
END_TRANSITION
TRANSITION FROM Ready TO R_Water
    := eProcess=E_CIP_Return.eT93_R_Water;
END_TRANSITION
STEP R_Water:
    _aR_Water_entry(P1);  // entry action
    _aR_Water_active(N);  // step action
END_STEP
TRANSITION FROM R_Water TO Done
    := bStepDone;
END_TRANSITION
TRANSITION FROM Ready TO Water
    := eProcess=E_CIP_Return.eT94_Water;
END_TRANSITION
STEP Water:
    _aWater_entry(P1);  // entry action
    _aWater_active(N);  // step action
END_STEP
TRANSITION FROM Water TO Done
    := bStepDone;
END_TRANSITION
STEP Done:  // min time T#0.2s
    _aDone_entry(P1);  // entry action
END_STEP
TRANSITION FROM Done TO Init
    := TRUE;
END_TRANSITION
// branch label Branch1_act_Oper
END_ACTION

ACTION act_Status:
IF bReady AND bDone OR TRUE THEN;
	IF TRUE 
	AND fbPis.m_CheckByRecipe(stPis:=stPis_Tank_Water, 			req:=E_Piston_Recipe_State.Release)
	AND fbPis.m_CheckByRecipe(stPis:=stPis_Tank_R_Water, 		req:=E_Piston_Recipe_State.Release)
	AND fbPis.m_CheckByRecipe(stPis:=stPis_Tank_Detergent, 		req:=E_Piston_Recipe_State.Release)
	AND fbPis.m_CheckByRecipe(stPis:=stPis_Tank_DisInfection, 	req:=E_Piston_Recipe_State.Release)
	AND fbPis.m_CheckByRecipe(stPis:=stPis_Drain, 				req:=E_Piston_Recipe_State.Release)
	AND fbPis.m_CheckByRecipe(stPis:=stPis_Tank_Water_1, 		req:=E_Piston_Recipe_State.Release)
	AND fbPis.m_CheckByRecipe(stPis:=stPis_Tank_R_Water_1, 		req:=E_Piston_Recipe_State.Release)
	AND fbPis.m_CheckByRecipe(stPis:=stPis_Tank_Detergent_1, 	req:=E_Piston_Recipe_State.Release)
	AND fbPis.m_CheckByRecipe(stPis:=stPis_Tank_DisInfection_1, req:=E_Piston_Recipe_State.Release)
	THEN;
		eStatus:=E_CIP_Return.eDrain;
	
	ELSIF TRUE 
	AND fbPis.m_CheckByRecipe(stPis:=stPis_Tank_Water, 			req:=E_Piston_Recipe_State.Act)
	AND fbPis.m_CheckByRecipe(stPis:=stPis_Tank_R_Water, 		req:=E_Piston_Recipe_State.Release)
	AND fbPis.m_CheckByRecipe(stPis:=stPis_Tank_Detergent, 		req:=E_Piston_Recipe_State.Release)
	AND fbPis.m_CheckByRecipe(stPis:=stPis_Tank_DisInfection, 	req:=E_Piston_Recipe_State.Release)
	AND fbPis.m_CheckByRecipe(stPis:=stPis_Drain, 				req:=E_Piston_Recipe_State.Act)
	AND fbPis.m_CheckByRecipe(stPis:=stPis_Tank_Water_1, 		req:=E_Piston_Recipe_State.Act)
	AND fbPis.m_CheckByRecipe(stPis:=stPis_Tank_R_Water_1, 		req:=E_Piston_Recipe_State.Release)
	AND fbPis.m_CheckByRecipe(stPis:=stPis_Tank_Detergent_1, 	req:=E_Piston_Recipe_State.Release)
	AND fbPis.m_CheckByRecipe(stPis:=stPis_Tank_DisInfection_1, req:=E_Piston_Recipe_State.Release)
	THEN;
		eStatus:=E_CIP_Return.eT94_Water;
		
	ELSIF TRUE 
	AND fbPis.m_CheckByRecipe(stPis:=stPis_Tank_Water, 			req:=E_Piston_Recipe_State.Release)
	AND fbPis.m_CheckByRecipe(stPis:=stPis_Tank_R_Water, 		req:=E_Piston_Recipe_State.Act)
	AND fbPis.m_CheckByRecipe(stPis:=stPis_Tank_Detergent, 		req:=E_Piston_Recipe_State.Release)
	AND fbPis.m_CheckByRecipe(stPis:=stPis_Tank_DisInfection, 	req:=E_Piston_Recipe_State.Release)
	AND fbPis.m_CheckByRecipe(stPis:=stPis_Drain, 				req:=E_Piston_Recipe_State.Release)
	AND fbPis.m_CheckByRecipe(stPis:=stPis_Tank_Water_1, 			req:=E_Piston_Recipe_State.Release)
	AND fbPis.m_CheckByRecipe(stPis:=stPis_Tank_R_Water_1, 			req:=E_Piston_Recipe_State.Act)
	AND fbPis.m_CheckByRecipe(stPis:=stPis_Tank_Detergent_1, 		req:=E_Piston_Recipe_State.Release)
	AND fbPis.m_CheckByRecipe(stPis:=stPis_Tank_DisInfection_1, 	req:=E_Piston_Recipe_State.Release)
	THEN;
		eStatus:=E_CIP_Return.eT93_R_Water;
		
	ELSIF TRUE 	
	AND fbPis.m_CheckByRecipe(stPis:=stPis_Tank_Water, 			req:=E_Piston_Recipe_State.Release)
	AND fbPis.m_CheckByRecipe(stPis:=stPis_Tank_R_Water, 		req:=E_Piston_Recipe_State.Release)
	AND fbPis.m_CheckByRecipe(stPis:=stPis_Tank_Detergent, 		req:=E_Piston_Recipe_State.Act)
	AND fbPis.m_CheckByRecipe(stPis:=stPis_Tank_DisInfection, 	req:=E_Piston_Recipe_State.Release)
	AND fbPis.m_CheckByRecipe(stPis:=stPis_Drain, 				req:=E_Piston_Recipe_State.Release)
	AND fbPis.m_CheckByRecipe(stPis:=stPis_Tank_Water_1, 			req:=E_Piston_Recipe_State.Release)
	AND fbPis.m_CheckByRecipe(stPis:=stPis_Tank_R_Water_1, 			req:=E_Piston_Recipe_State.Release)
	AND fbPis.m_CheckByRecipe(stPis:=stPis_Tank_Detergent_1, 		req:=E_Piston_Recipe_State.Act)
	AND fbPis.m_CheckByRecipe(stPis:=stPis_Tank_DisInfection_1, 	req:=E_Piston_Recipe_State.Release)
	THEN;
		eStatus:=E_CIP_Return.eT92_Detergent;
		
	ELSIF TRUE 	
	AND fbPis.m_CheckByRecipe(stPis:=stPis_Tank_Water, 			req:=E_Piston_Recipe_State.Release)
	AND fbPis.m_CheckByRecipe(stPis:=stPis_Tank_R_Water, 		req:=E_Piston_Recipe_State.Release)
	AND fbPis.m_CheckByRecipe(stPis:=stPis_Tank_Detergent, 		req:=E_Piston_Recipe_State.Release)
	AND fbPis.m_CheckByRecipe(stPis:=stPis_Tank_DisInfection, 	req:=E_Piston_Recipe_State.Act)
	AND fbPis.m_CheckByRecipe(stPis:=stPis_Drain, 				req:=E_Piston_Recipe_State.Release)
	AND fbPis.m_CheckByRecipe(stPis:=stPis_Tank_Water_1, 			req:=E_Piston_Recipe_State.Release)
	AND fbPis.m_CheckByRecipe(stPis:=stPis_Tank_R_Water_1, 			req:=E_Piston_Recipe_State.Release)
	AND fbPis.m_CheckByRecipe(stPis:=stPis_Tank_Detergent_1, 		req:=E_Piston_Recipe_State.Release)
	AND fbPis.m_CheckByRecipe(stPis:=stPis_Tank_DisInfection_1, 	req:=E_Piston_Recipe_State.Act)
	THEN;
		eStatus:=E_CIP_Return.eT91_Sanitation;
	ELSE;
		eStatus:=E_CIP_Return.eNone;
	END_IF
ELSE;
	eStatus:=E_CIP_Return.eNone;
END_IF
END_ACTION

METHOD m_CheckStatus : BOOL
VAR_INPUT
	eReqStatus		: E_CIP_Return;
END_VAR
IF eStatus=eReqStatus 
AND eProcess=E_CIP_Return.eNone
AND eReq=E_CIP_Return.eNone
AND bReady
AND bDone
AND NOT bRun
THEN;
	m_CheckStatus:=TRUE;
END_IF
END_METHOD

METHOD m_Request_Reset : BOOL
VAR_IN_OUT
	memo: R_TRIG;
END_VAR
memo(CLK:=eReq=0);
IF TRUE 
AND memo.Q
THEN;
	SFCReset:=TRUE;
END_IF
END_METHOD

METHOD m_Run : BOOL
VAR_INPUT
	eReqProc			: E_CIP_Return;
END_VAR
IF eProcess=E_CIP_Return.eNone THEN;
	eProcess:=eReq:=eReqProc;
	bDone:=FALSE;
	m_Run:=TRUE;
END_IF
END_METHOD

METHOD m_Set_SFCFlags_Reference : BOOL
//Set reference to SFC flags

refSFC.SFCInit REF= SFCInit;
refSFC.SFCReset REF= SFCReset;
refSFC.SFCError REF= SFCError;
refSFC.SFCEnableLimit REF= SFCEnableLimit;
refSFC.SFCErrorStep REF= SFCErrorStep;
refSFC.SFCErrorPOU REF= SFCErrorPOU;
refSFC.SFCQuitError REF= SFCQuitError;
refSFC.SFCPause REF= SFCPause;
refSFC.SFCTrans REF= SFCTrans;
refSFC.SFCCurrentStep REF= SFCCurrentStep;
refSFC.SFCTip REF= SFCTip;
refSFC.SFCTipMode REF= SFCTipMode;

// Cycle handle for SFC
m_SFC_Handle();
END_METHOD

END_FUNCTION_BLOCK

// ---- 03 Project/23 CIP/FB_CIP_Client.TcPOU
FUNCTION_BLOCK FB_CIP_Client EXTENDS FB_SFC_Cycle IMPLEMENTS ITF_FB_SFC_Cycle
VAR_INPUT
	//eElementID			: E_Element_List;
	
	valClient_Source		: E_Pis_Name;
	valClient_Return		: E_Pis_Name;
	valS_Marinade_Up		: E_Pis_Name;
	//valS_Marinade_Up_Drain	: E_Pis_Name;
	valS_Marinade_Low		: E_Pis_Name;
	valS_Color_Up			: E_Pis_Name;
	//valS_Color_Up_Drain		: E_Pis_Name;
	valS_Color_Low			: E_Pis_Name;
	//valTank_1				: E_Pis_Name;
	//valTank_2				: E_Pis_Name;
	//valTank_3				: E_Pis_Name;
	//valTank_4				: E_Pis_Name;
	//valS_Marinade_Low_Select	: E_Pis_Name;
	//valS_Color_Low_Select	: E_Pis_Name;
	valDrain				: E_Pis_Name;
	valLoop					: E_Pis_Name;//V1030
	valS_Future				: E_Pis_Name;
	
END_VAR
VAR_OUTPUT
END_VAR
VAR
	//refElement		: REFERENCE TO FB_Element;
	//refState_Long		: REFERENCE TO E_Element_State_Long;
	eReq				: E_CIP_Client_Selector;
	eProcess			: E_CIP_Client_Selector;
	eStatus				: E_CIP_Client_Selector;
	
	fbPis					: FB_Piston;
	stPis_Client_Source			: REFERENCE TO ST_Piston;
	stPis_Client_Return			: REFERENCE TO ST_Piston;
	stPis_S_Marinade_Up			: REFERENCE TO ST_Piston;
	//stPis_S_Marinade_Up_Drain	: REFERENCE TO ST_Piston;
	stPis_S_Marinade_Low		: REFERENCE TO ST_Piston;
	stPis_S_Color_Up			: REFERENCE TO ST_Piston;
	//stPis_S_Color_Up_Drain		: REFERENCE TO ST_Piston;
	stPis_S_Color_Low			: REFERENCE TO ST_Piston;
	//stPis_Tank_1				: REFERENCE TO ST_Piston;
	//stPis_Tank_2				: REFERENCE TO ST_Piston;
	//stPis_Tank_3				: REFERENCE TO ST_Piston;
	//stPis_Tank_4				: REFERENCE TO ST_Piston;
	//stPis_S_Marinade_Low_Select	: REFERENCE TO ST_Piston;
	//stPis_S_Color_Low_Select	: REFERENCE TO ST_Piston;
	stPis_Drain					: REFERENCE TO ST_Piston;	
	stPis_Loop					: REFERENCE TO ST_Piston;//V1030
	stPis_S_Future				: REFERENCE TO ST_Piston;

	tonDrainTime: TON;
	
	rt_Req_Reset: R_TRIG;

END_VAR
VAR_IN_OUT


END_VAR

act_GetReference();

act_Oper();
IF NOT Init.x THEN;
	act_Status();
END_IF

tonDrainTime(PT:=T#1M, IN:=eStatus=E_CIP_Client_Selector.eDrain);
IF tonDrainTime.Q 
AND eReq=E_CIP_Client_Selector.eNone
AND eProcess=E_CIP_Client_Selector.eNone
THEN;
	eReq:=E_CIP_Client_Selector.eClose;
END_IF

m_Request_Reset(memo:=rt_Req_Reset);//rt_Req_Reset: R_TRIG;

ACTION _aClose_active:
bStepDone:=FALSE;
IF TRUE 
AND eStatus=E_CIP_Client_Selector.eClose
THEN;
	bStepDone:=TRUE;
END_IF
END_ACTION

ACTION _aClose_entry:
fbPis.m_SetByRecipe(stPis:=stPis_Client_Source, 		req:=E_Piston_Recipe_State.Release);
fbPis.m_SetByRecipe(stPis:=stPis_Client_Return, 		req:=E_Piston_Recipe_State.Release);
fbPis.m_SetByRecipe(stPis:=stPis_S_Marinade_Up, 		req:=E_Piston_Recipe_State.Release);
fbPis.m_SetByRecipe(stPis:=stPis_S_Marinade_Low, 		req:=E_Piston_Recipe_State.Release);
fbPis.m_SetByRecipe(stPis:=stPis_S_Color_Up, 			req:=E_Piston_Recipe_State.Release);
fbPis.m_SetByRecipe(stPis:=stPis_S_Color_Low, 			req:=E_Piston_Recipe_State.Release);
fbPis.m_SetByRecipe(stPis:=stPis_Drain, 				req:=E_Piston_Recipe_State.Release);
fbPis.m_SetByRecipe(stPis:=stPis_Loop, 					req:=E_Piston_Recipe_State.Release);
fbPis.m_SetByRecipe(stPis:=stPis_S_Future, 				req:=E_Piston_Recipe_State.Release);
END_ACTION

ACTION _aColor_Low_active:
bStepDone:=FALSE;
IF TRUE 
AND eStatus=E_CIP_Client_Selector.eColor_Low
THEN;
	bStepDone:=TRUE;
END_IF
END_ACTION

ACTION _aColor_Low_entry:
fbPis.m_SetByRecipe(stPis:=stPis_Client_Source, 		req:=E_Piston_Recipe_State.Act);
fbPis.m_SetByRecipe(stPis:=stPis_Client_Return, 		req:=E_Piston_Recipe_State.Act);
fbPis.m_SetByRecipe(stPis:=stPis_S_Marinade_Up, 		req:=E_Piston_Recipe_State.Release);
fbPis.m_SetByRecipe(stPis:=stPis_S_Marinade_Low, 		req:=E_Piston_Recipe_State.Release);
fbPis.m_SetByRecipe(stPis:=stPis_S_Color_Up, 			req:=E_Piston_Recipe_State.Release);
fbPis.m_SetByRecipe(stPis:=stPis_S_Color_Low, 			req:=E_Piston_Recipe_State.Act);
fbPis.m_SetByRecipe(stPis:=stPis_Drain, 				req:=E_Piston_Recipe_State.Release);
fbPis.m_SetByRecipe(stPis:=stPis_Loop, 					req:=E_Piston_Recipe_State.Release);
fbPis.m_SetByRecipe(stPis:=stPis_S_Future, 				req:=E_Piston_Recipe_State.Release);
END_ACTION

ACTION _aColor_Up_active:
bStepDone:=FALSE;
IF TRUE 
AND eStatus=E_CIP_Client_Selector.eColor_Up
THEN;
	bStepDone:=TRUE;
END_IF
END_ACTION

ACTION _aColor_Up_entry:
fbPis.m_SetByRecipe(stPis:=stPis_Client_Source, 		req:=E_Piston_Recipe_State.Act);
fbPis.m_SetByRecipe(stPis:=stPis_Client_Return, 		req:=E_Piston_Recipe_State.Act);
fbPis.m_SetByRecipe(stPis:=stPis_S_Marinade_Up, 		req:=E_Piston_Recipe_State.Release);
fbPis.m_SetByRecipe(stPis:=stPis_S_Marinade_Low, 		req:=E_Piston_Recipe_State.Release);
fbPis.m_SetByRecipe(stPis:=stPis_S_Color_Up, 			req:=E_Piston_Recipe_State.Act);
fbPis.m_SetByRecipe(stPis:=stPis_S_Color_Low, 			req:=E_Piston_Recipe_State.Release);
fbPis.m_SetByRecipe(stPis:=stPis_Drain, 				req:=E_Piston_Recipe_State.Release);
fbPis.m_SetByRecipe(stPis:=stPis_Loop, 					req:=E_Piston_Recipe_State.Release);
fbPis.m_SetByRecipe(stPis:=stPis_S_Future, 				req:=E_Piston_Recipe_State.Release);
END_ACTION

ACTION _aDone_entry:
eProcess:=E_CIP_Usage.eNotInUse;
eReq:=E_CIP_Usage.eNotInUse;
bRun:=FALSE;
bDone:=TRUE;
END_ACTION

ACTION _aDrain_active:
bStepDone:=FALSE;
IF TRUE 
AND eStatus=E_CIP_Client_Selector.eDrain
THEN;
	bStepDone:=TRUE;
END_IF
END_ACTION

ACTION _aDrain_entry:
fbPis.m_SetByRecipe(stPis:=stPis_Client_Source, 		req:=E_Piston_Recipe_State.Release);
fbPis.m_SetByRecipe(stPis:=stPis_Client_Return, 		req:=E_Piston_Recipe_State.Release);
fbPis.m_SetByRecipe(stPis:=stPis_S_Marinade_Up, 		req:=E_Piston_Recipe_State.Release);
fbPis.m_SetByRecipe(stPis:=stPis_S_Marinade_Low, 		req:=E_Piston_Recipe_State.Release);
fbPis.m_SetByRecipe(stPis:=stPis_S_Color_Up, 			req:=E_Piston_Recipe_State.Release);
fbPis.m_SetByRecipe(stPis:=stPis_S_Color_Low, 			req:=E_Piston_Recipe_State.Release);
fbPis.m_SetByRecipe(stPis:=stPis_Drain, 				req:=E_Piston_Recipe_State.Act);
fbPis.m_SetByRecipe(stPis:=stPis_Loop, 					req:=E_Piston_Recipe_State.Release);
fbPis.m_SetByRecipe(stPis:=stPis_S_Future, 				req:=E_Piston_Recipe_State.Release);
END_ACTION

ACTION _aFuture_active:
bStepDone:=FALSE;
IF TRUE 
AND eStatus=E_CIP_Client_Selector.eFuture
THEN;
	bStepDone:=TRUE;
END_IF
END_ACTION

ACTION _aFuture_entry:
fbPis.m_SetByRecipe(stPis:=stPis_Client_Source, 		req:=E_Piston_Recipe_State.Act);
fbPis.m_SetByRecipe(stPis:=stPis_Client_Return, 		req:=E_Piston_Recipe_State.Act);
fbPis.m_SetByRecipe(stPis:=stPis_S_Marinade_Up, 		req:=E_Piston_Recipe_State.Release);
fbPis.m_SetByRecipe(stPis:=stPis_S_Marinade_Low, 		req:=E_Piston_Recipe_State.Release);
fbPis.m_SetByRecipe(stPis:=stPis_S_Color_Up, 			req:=E_Piston_Recipe_State.Release);
fbPis.m_SetByRecipe(stPis:=stPis_S_Color_Low, 			req:=E_Piston_Recipe_State.Release);
fbPis.m_SetByRecipe(stPis:=stPis_Drain, 				req:=E_Piston_Recipe_State.Release);
fbPis.m_SetByRecipe(stPis:=stPis_Loop, 					req:=E_Piston_Recipe_State.Release);
fbPis.m_SetByRecipe(stPis:=stPis_S_Future, 				req:=E_Piston_Recipe_State.Act);
END_ACTION

ACTION _aInit_active:
SFCReset:=FALSE;
END_ACTION

ACTION _aInit_exit:
eProcess:=E_CIP_Usage.eNotInUse;
eReq:=E_CIP_Usage.eNotInUse;
END_ACTION

ACTION _aLoop_active:
bStepDone:=FALSE;
IF TRUE 
AND eStatus=E_CIP_Client_Selector.eLoop
THEN;
	bStepDone:=TRUE;
END_IF
END_ACTION

ACTION _aLoop_entry:
fbPis.m_SetByRecipe(stPis:=stPis_Client_Source, 		req:=E_Piston_Recipe_State.Act);
fbPis.m_SetByRecipe(stPis:=stPis_Client_Return, 		req:=E_Piston_Recipe_State.Act);
fbPis.m_SetByRecipe(stPis:=stPis_S_Marinade_Up, 		req:=E_Piston_Recipe_State.Release);
fbPis.m_SetByRecipe(stPis:=stPis_S_Marinade_Low, 		req:=E_Piston_Recipe_State.Release);
fbPis.m_SetByRecipe(stPis:=stPis_S_Color_Up, 			req:=E_Piston_Recipe_State.Release);
fbPis.m_SetByRecipe(stPis:=stPis_S_Color_Low, 			req:=E_Piston_Recipe_State.Release);
fbPis.m_SetByRecipe(stPis:=stPis_Drain, 				req:=E_Piston_Recipe_State.Act);
fbPis.m_SetByRecipe(stPis:=stPis_Loop, 					req:=E_Piston_Recipe_State.Act);
fbPis.m_SetByRecipe(stPis:=stPis_S_Future, 				req:=E_Piston_Recipe_State.Release);
END_ACTION

ACTION _aMarinade_Low_active:
bStepDone:=FALSE;
IF TRUE 
AND eStatus=E_CIP_Client_Selector.eMarinade_Low
THEN;
	bStepDone:=TRUE;
END_IF
END_ACTION

ACTION _aMarinade_Low_entry:
fbPis.m_SetByRecipe(stPis:=stPis_Client_Source, 		req:=E_Piston_Recipe_State.Act);
fbPis.m_SetByRecipe(stPis:=stPis_Client_Return, 		req:=E_Piston_Recipe_State.Act);
fbPis.m_SetByRecipe(stPis:=stPis_S_Marinade_Up, 		req:=E_Piston_Recipe_State.Release);
fbPis.m_SetByRecipe(stPis:=stPis_S_Marinade_Low, 		req:=E_Piston_Recipe_State.Act);
fbPis.m_SetByRecipe(stPis:=stPis_S_Color_Up, 			req:=E_Piston_Recipe_State.Release);
fbPis.m_SetByRecipe(stPis:=stPis_S_Color_Low, 			req:=E_Piston_Recipe_State.Release);
fbPis.m_SetByRecipe(stPis:=stPis_Drain, 				req:=E_Piston_Recipe_State.Release);
fbPis.m_SetByRecipe(stPis:=stPis_Loop, 					req:=E_Piston_Recipe_State.Release);
fbPis.m_SetByRecipe(stPis:=stPis_S_Future, 				req:=E_Piston_Recipe_State.Release);
END_ACTION

ACTION _aMarinade_Up_active:
bStepDone:=FALSE;
IF TRUE 
AND eStatus=E_CIP_Client_Selector.eMarinade_Up
THEN;
	bStepDone:=TRUE;
END_IF
END_ACTION

ACTION _aMarinade_Up_entry:
fbPis.m_SetByRecipe(stPis:=stPis_Client_Source, 		req:=E_Piston_Recipe_State.Act);
fbPis.m_SetByRecipe(stPis:=stPis_Client_Return, 		req:=E_Piston_Recipe_State.Act);
fbPis.m_SetByRecipe(stPis:=stPis_S_Marinade_Up, 		req:=E_Piston_Recipe_State.Act);
fbPis.m_SetByRecipe(stPis:=stPis_S_Marinade_Low, 		req:=E_Piston_Recipe_State.Release);
fbPis.m_SetByRecipe(stPis:=stPis_S_Color_Up, 			req:=E_Piston_Recipe_State.Release);
fbPis.m_SetByRecipe(stPis:=stPis_S_Color_Low, 			req:=E_Piston_Recipe_State.Release);
fbPis.m_SetByRecipe(stPis:=stPis_Drain, 				req:=E_Piston_Recipe_State.Release);
fbPis.m_SetByRecipe(stPis:=stPis_Loop, 					req:=E_Piston_Recipe_State.Release);
fbPis.m_SetByRecipe(stPis:=stPis_S_Future, 				req:=E_Piston_Recipe_State.Release);
END_ACTION

ACTION _aReady_active:


IF eReq<>E_CIP_Client_Selector.eNone THEN;
	IF eProcess=E_CIP_Client_Selector.eNone 
	THEN;
		eProcess:=eReq;
	ELSE;
		eReq:=E_CIP_Client_Selector.eNone;
	END_IF
END_IF

(*
CASE eReq OF
	E_CIP_Usage.eLine_Color:;
			IF TRUE THEN;
				eProcess:=E_CIP_Usage.eLine_Color;
			END_IF

	E_CIP_Usage.eLine_Marinada:;
			IF TRUE THEN;
				eProcess:=E_CIP_Usage.eLine_Marinada;
			END_IF	
			
	E_CIP_Usage.eLocal:;
			IF TRUE THEN;
				eProcess:=E_CIP_Usage.eLocal;
			END_IF	

	E_CIP_Usage.eNotInUse:;
			IF TRUE THEN;
				eProcess:=E_CIP_Usage.eNotInUse;
			END_IF	
			
	E_CIP_Usage.eTank_1:;
			IF TRUE THEN;
				eProcess:=E_CIP_Usage.eTank_1;
			END_IF	
	E_CIP_Usage.eTank_2:;
			IF TRUE THEN;
				eProcess:=E_CIP_Usage.eTank_2;
			END_IF	
	E_CIP_Usage.eTank_3:;
			IF TRUE THEN;
				eProcess:=E_CIP_Usage.eTank_3;
			END_IF	
	E_CIP_Usage.eTank_4:;
			IF TRUE THEN;
				eProcess:=E_CIP_Usage.eTank_4;
			END_IF	
	E_CIP_Usage.eTriBlender_Color:;
			IF TRUE THEN;
				eProcess:=E_CIP_Usage.eTriBlender_Color;
			END_IF	
	E_CIP_Usage.eTriBlender_Marinada:;
			IF TRUE THEN;
				eProcess:=E_CIP_Usage.eTriBlender_Marinada;
			END_IF	

END_CASE
*)
END_ACTION

ACTION _aReady_exit:
bRun:=TRUE;
bDone:=FALSE;
END_ACTION

ACTION act_GetReference:
m_Set_SFCFlags_Reference();
//refElement REF= fbElement[eElementID];
//refState_Long REF= fbElement[eElementID].eState_Long;

stPis_Client_Source			REF= g_Piston.stPis[valClient_Source];
stPis_Client_Return			REF= g_Piston.stPis[valClient_Return];
stPis_S_Marinade_Up			REF= g_Piston.stPis[valS_Marinade_Up];
//stPis_S_Marinade_Up_Drain	REF= g_Piston.stPis[valS_Marinade_Up_Drain];
stPis_S_Marinade_Low		REF= g_Piston.stPis[valS_Marinade_Low];
stPis_S_Color_Up			REF= g_Piston.stPis[valS_Color_Up];
//stPis_S_Color_Up_Drain		REF= g_Piston.stPis[valS_Color_Up_Drain];
stPis_S_Color_Low			REF= g_Piston.stPis[valS_Color_Low];
//stPis_Tank_1				REF= g_Piston.stPis[valTank_1];
//stPis_Tank_2				REF= g_Piston.stPis[valTank_2];
//stPis_Tank_3				REF= g_Piston.stPis[valTank_3];
//stPis_Tank_4				REF= g_Piston.stPis[valTank_4];
//stPis_S_Marinade_Low_Select	REF= g_Piston.stPis[valS_Marinade_Low_Select];
//stPis_S_Color_Low_Select	REF= g_Piston.stPis[valS_Color_Low_Select];
stPis_Drain					REF= g_Piston.stPis[valDrain];
stPis_Loop				REF= g_Piston.stPis[valLoop];
stPis_S_Future				REF= g_Piston.stPis[valS_Future];
END_ACTION

ACTION act_Oper:
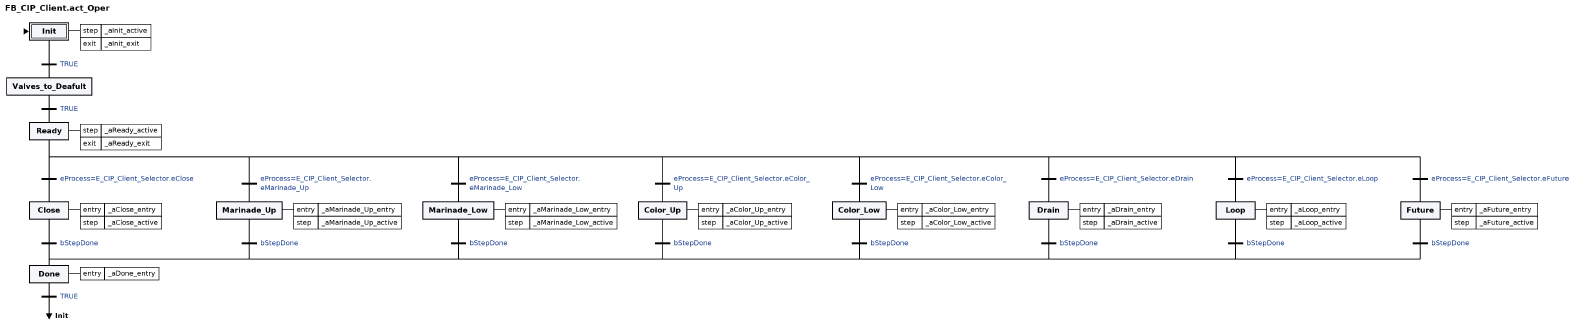
INITIAL_STEP Init:  // min time T#0.5s
    _aInit_active(N);  // step action
    _aInit_exit(P0);  // exit action
END_STEP
TRANSITION FROM Init TO Valves_to_Deafult
    := TRUE;
END_TRANSITION
STEP Valves_to_Deafult:
END_STEP
TRANSITION FROM Valves_to_Deafult TO Ready
    := TRUE;
END_TRANSITION
STEP Ready:
    _aReady_active(N);  // step action
    _aReady_exit(P0);  // exit action
END_STEP
TRANSITION FROM Ready TO Close
    := eProcess=E_CIP_Client_Selector.eClose;
END_TRANSITION
STEP Close:
    _aClose_entry(P1);  // entry action
    _aClose_active(N);  // step action
END_STEP
TRANSITION FROM Close TO Done
    := bStepDone;
END_TRANSITION
TRANSITION FROM Ready TO Marinade_Up
    := eProcess=E_CIP_Client_Selector.eMarinade_Up;
END_TRANSITION
STEP Marinade_Up:
    _aMarinade_Up_entry(P1);  // entry action
    _aMarinade_Up_active(N);  // step action
END_STEP
TRANSITION FROM Marinade_Up TO Done
    := bStepDone;
END_TRANSITION
TRANSITION FROM Ready TO Marinade_Low
    := eProcess=E_CIP_Client_Selector.eMarinade_Low;
END_TRANSITION
STEP Marinade_Low:
    _aMarinade_Low_entry(P1);  // entry action
    _aMarinade_Low_active(N);  // step action
END_STEP
TRANSITION FROM Marinade_Low TO Done
    := bStepDone;
END_TRANSITION
TRANSITION FROM Ready TO Color_Up
    := eProcess=E_CIP_Client_Selector.eColor_Up;
END_TRANSITION
STEP Color_Up:
    _aColor_Up_entry(P1);  // entry action
    _aColor_Up_active(N);  // step action
END_STEP
TRANSITION FROM Color_Up TO Done
    := bStepDone;
END_TRANSITION
TRANSITION FROM Ready TO Color_Low
    := eProcess=E_CIP_Client_Selector.eColor_Low;
END_TRANSITION
STEP Color_Low:
    _aColor_Low_entry(P1);  // entry action
    _aColor_Low_active(N);  // step action
END_STEP
TRANSITION FROM Color_Low TO Done
    := bStepDone;
END_TRANSITION
TRANSITION FROM Ready TO Drain
    := eProcess=E_CIP_Client_Selector.eDrain;
END_TRANSITION
STEP Drain:
    _aDrain_entry(P1);  // entry action
    _aDrain_active(N);  // step action
END_STEP
TRANSITION FROM Drain TO Done
    := bStepDone;
END_TRANSITION
TRANSITION FROM Ready TO Loop
    := eProcess=E_CIP_Client_Selector.eLoop;
END_TRANSITION
STEP Loop:
    _aLoop_entry(P1);  // entry action
    _aLoop_active(N);  // step action
END_STEP
TRANSITION FROM Loop TO Done
    := bStepDone;
END_TRANSITION
TRANSITION FROM Ready TO Future
    := eProcess=E_CIP_Client_Selector.eFuture;
END_TRANSITION
STEP Future:
    _aFuture_entry(P1);  // entry action
    _aFuture_active(N);  // step action
END_STEP
TRANSITION FROM Future TO Done
    := bStepDone;
END_TRANSITION
STEP Done:  // min time T#0.2s
    _aDone_entry(P1);  // entry action
END_STEP
TRANSITION FROM Done TO Init
    := TRUE;
END_TRANSITION
// branch label Branch2_act_Oper
END_ACTION

ACTION act_Status:
IF bReady AND bDone OR TRUE THEN;
	IF TRUE 
	AND fbPis.m_CheckByRecipe(stPis:=stPis_Client_Source, 		req:=E_Piston_Recipe_State.Release)
	AND fbPis.m_CheckByRecipe(stPis:=stPis_Client_Return, 		req:=E_Piston_Recipe_State.Release)
	AND fbPis.m_CheckByRecipe(stPis:=stPis_S_Marinade_Up, 		req:=E_Piston_Recipe_State.Release)
	AND fbPis.m_CheckByRecipe(stPis:=stPis_S_Marinade_Low, 		req:=E_Piston_Recipe_State.Release)
	AND fbPis.m_CheckByRecipe(stPis:=stPis_S_Color_Up, 			req:=E_Piston_Recipe_State.Release)
	AND fbPis.m_CheckByRecipe(stPis:=stPis_S_Color_Low, 		req:=E_Piston_Recipe_State.Release)
	AND fbPis.m_CheckByRecipe(stPis:=stPis_Drain, 				req:=E_Piston_Recipe_State.Release)
	AND fbPis.m_CheckByRecipe(stPis:=stPis_Loop, 				req:=E_Piston_Recipe_State.Release)
	AND fbPis.m_CheckByRecipe(stPis:=stPis_S_Future, 			req:=E_Piston_Recipe_State.Release)
	THEN;
		eStatus:=E_CIP_Client_Selector.eClose;
	ELSIF TRUE
	AND fbPis.m_CheckByRecipe(stPis:=stPis_Client_Source, 		req:=E_Piston_Recipe_State.Act)
	AND fbPis.m_CheckByRecipe(stPis:=stPis_Client_Return, 		req:=E_Piston_Recipe_State.Act)
	AND fbPis.m_CheckByRecipe(stPis:=stPis_S_Marinade_Up, 		req:=E_Piston_Recipe_State.Act)
	AND fbPis.m_CheckByRecipe(stPis:=stPis_S_Marinade_Low, 		req:=E_Piston_Recipe_State.Release)
	AND fbPis.m_CheckByRecipe(stPis:=stPis_S_Color_Up, 			req:=E_Piston_Recipe_State.Release)
	AND fbPis.m_CheckByRecipe(stPis:=stPis_S_Color_Low, 		req:=E_Piston_Recipe_State.Release)
	AND fbPis.m_CheckByRecipe(stPis:=stPis_Drain, 				req:=E_Piston_Recipe_State.Release)
	AND fbPis.m_CheckByRecipe(stPis:=stPis_Loop, 				req:=E_Piston_Recipe_State.Release)
	AND fbPis.m_CheckByRecipe(stPis:=stPis_S_Future, 			req:=E_Piston_Recipe_State.Release)
	THEN;
		eStatus:=E_CIP_Client_Selector.eMarinade_Up;
	ELSIF TRUE 
	AND fbPis.m_CheckByRecipe(stPis:=stPis_Client_Source, 		req:=E_Piston_Recipe_State.Act)
	AND fbPis.m_CheckByRecipe(stPis:=stPis_Client_Return, 		req:=E_Piston_Recipe_State.Act)
	AND fbPis.m_CheckByRecipe(stPis:=stPis_S_Marinade_Up, 		req:=E_Piston_Recipe_State.Release)
	AND fbPis.m_CheckByRecipe(stPis:=stPis_S_Marinade_Low, 		req:=E_Piston_Recipe_State.Act)
	AND fbPis.m_CheckByRecipe(stPis:=stPis_S_Color_Up, 			req:=E_Piston_Recipe_State.Release)
	AND fbPis.m_CheckByRecipe(stPis:=stPis_S_Color_Low, 		req:=E_Piston_Recipe_State.Release)
	AND fbPis.m_CheckByRecipe(stPis:=stPis_Drain, 				req:=E_Piston_Recipe_State.Release)
	AND fbPis.m_CheckByRecipe(stPis:=stPis_Loop, 				req:=E_Piston_Recipe_State.Release)
	AND fbPis.m_CheckByRecipe(stPis:=stPis_S_Future, 			req:=E_Piston_Recipe_State.Release)
	THEN;
		eStatus:=E_CIP_Client_Selector.eMarinade_Low;
	ELSIF TRUE 
	AND fbPis.m_CheckByRecipe(stPis:=stPis_Client_Source, 		req:=E_Piston_Recipe_State.Act)
	AND fbPis.m_CheckByRecipe(stPis:=stPis_Client_Return, 		req:=E_Piston_Recipe_State.Act)
	AND fbPis.m_CheckByRecipe(stPis:=stPis_S_Marinade_Up, 		req:=E_Piston_Recipe_State.Release)
	AND fbPis.m_CheckByRecipe(stPis:=stPis_S_Marinade_Low, 		req:=E_Piston_Recipe_State.Release)
	AND fbPis.m_CheckByRecipe(stPis:=stPis_S_Color_Up, 			req:=E_Piston_Recipe_State.Act)
	AND fbPis.m_CheckByRecipe(stPis:=stPis_S_Color_Low, 		req:=E_Piston_Recipe_State.Release)
	AND fbPis.m_CheckByRecipe(stPis:=stPis_Drain, 				req:=E_Piston_Recipe_State.Release)
	AND fbPis.m_CheckByRecipe(stPis:=stPis_Loop, 				req:=E_Piston_Recipe_State.Release)
	AND fbPis.m_CheckByRecipe(stPis:=stPis_S_Future, 			req:=E_Piston_Recipe_State.Release)
	THEN;
		eStatus:=E_CIP_Client_Selector.eColor_Up;
	ELSIF TRUE 
	AND fbPis.m_CheckByRecipe(stPis:=stPis_Client_Source, 		req:=E_Piston_Recipe_State.Act)
	AND fbPis.m_CheckByRecipe(stPis:=stPis_Client_Return, 		req:=E_Piston_Recipe_State.Act)
	AND fbPis.m_CheckByRecipe(stPis:=stPis_S_Marinade_Up, 		req:=E_Piston_Recipe_State.Release)
	AND fbPis.m_CheckByRecipe(stPis:=stPis_S_Marinade_Low, 		req:=E_Piston_Recipe_State.Release)
	AND fbPis.m_CheckByRecipe(stPis:=stPis_S_Color_Up, 			req:=E_Piston_Recipe_State.Release)
	AND fbPis.m_CheckByRecipe(stPis:=stPis_S_Color_Low, 		req:=E_Piston_Recipe_State.Act)
	AND fbPis.m_CheckByRecipe(stPis:=stPis_Drain, 				req:=E_Piston_Recipe_State.Release)
	AND fbPis.m_CheckByRecipe(stPis:=stPis_Loop, 				req:=E_Piston_Recipe_State.Release)
	AND fbPis.m_CheckByRecipe(stPis:=stPis_S_Future, 			req:=E_Piston_Recipe_State.Release)
	THEN;
		eStatus:=E_CIP_Client_Selector.eColor_Low;
	ELSIF TRUE 
	AND fbPis.m_CheckByRecipe(stPis:=stPis_Client_Source, 		req:=E_Piston_Recipe_State.Release)
	AND fbPis.m_CheckByRecipe(stPis:=stPis_Client_Return, 		req:=E_Piston_Recipe_State.Release)
	AND fbPis.m_CheckByRecipe(stPis:=stPis_S_Marinade_Up, 		req:=E_Piston_Recipe_State.Release)
	AND fbPis.m_CheckByRecipe(stPis:=stPis_S_Marinade_Low, 		req:=E_Piston_Recipe_State.Release)
	AND fbPis.m_CheckByRecipe(stPis:=stPis_S_Color_Up, 			req:=E_Piston_Recipe_State.Release)
	AND fbPis.m_CheckByRecipe(stPis:=stPis_S_Color_Low, 		req:=E_Piston_Recipe_State.Release)
	AND fbPis.m_CheckByRecipe(stPis:=stPis_Drain, 				req:=E_Piston_Recipe_State.Act)
	AND fbPis.m_CheckByRecipe(stPis:=stPis_Loop, 				req:=E_Piston_Recipe_State.Release)
	AND fbPis.m_CheckByRecipe(stPis:=stPis_S_Future, 			req:=E_Piston_Recipe_State.Release)
	THEN;
		eStatus:=E_CIP_Client_Selector.eDrain;
	ELSIF TRUE 
	AND fbPis.m_CheckByRecipe(stPis:=stPis_Client_Source, 		req:=E_Piston_Recipe_State.Act)
	AND fbPis.m_CheckByRecipe(stPis:=stPis_Client_Return, 		req:=E_Piston_Recipe_State.Act)
	AND fbPis.m_CheckByRecipe(stPis:=stPis_S_Marinade_Up, 		req:=E_Piston_Recipe_State.Release)
	AND fbPis.m_CheckByRecipe(stPis:=stPis_S_Marinade_Low, 		req:=E_Piston_Recipe_State.Release)
	AND fbPis.m_CheckByRecipe(stPis:=stPis_S_Color_Up, 			req:=E_Piston_Recipe_State.Release)
	AND fbPis.m_CheckByRecipe(stPis:=stPis_S_Color_Low, 		req:=E_Piston_Recipe_State.Release)
	AND fbPis.m_CheckByRecipe(stPis:=stPis_Drain, 				req:=E_Piston_Recipe_State.Act)
	AND fbPis.m_CheckByRecipe(stPis:=stPis_Loop, 				req:=E_Piston_Recipe_State.Act)
	AND fbPis.m_CheckByRecipe(stPis:=stPis_S_Future, 			req:=E_Piston_Recipe_State.Release)
	THEN;
		eStatus:=E_CIP_Client_Selector.eLoop;
	ELSIF TRUE 
	AND fbPis.m_CheckByRecipe(stPis:=stPis_Client_Source, 		req:=E_Piston_Recipe_State.Act)
	AND fbPis.m_CheckByRecipe(stPis:=stPis_Client_Return, 		req:=E_Piston_Recipe_State.Act)
	AND fbPis.m_CheckByRecipe(stPis:=stPis_S_Marinade_Up, 		req:=E_Piston_Recipe_State.Release)
	AND fbPis.m_CheckByRecipe(stPis:=stPis_S_Marinade_Low, 		req:=E_Piston_Recipe_State.Release)
	AND fbPis.m_CheckByRecipe(stPis:=stPis_S_Color_Up, 			req:=E_Piston_Recipe_State.Release)
	AND fbPis.m_CheckByRecipe(stPis:=stPis_S_Color_Low, 		req:=E_Piston_Recipe_State.Release)
	AND fbPis.m_CheckByRecipe(stPis:=stPis_Drain, 				req:=E_Piston_Recipe_State.Release)
	AND fbPis.m_CheckByRecipe(stPis:=stPis_Loop, 				req:=E_Piston_Recipe_State.Release)
	AND fbPis.m_CheckByRecipe(stPis:=stPis_S_Future, 			req:=E_Piston_Recipe_State.Act)
	THEN;
		eStatus:=E_CIP_Client_Selector.eFuture;
	ELSE;
		eStatus:=E_CIP_Client_Selector.eNone;
	END_IF
ELSE;
	eStatus:=E_CIP_Client_Selector.eNone;
END_IF
END_ACTION

METHOD m_CheckStatus : BOOL
VAR_INPUT
	eReqStatus		: E_CIP_Usage;
END_VAR
VAR
	eReqStatusLocal	: E_CIP_Client_Selector;
END_VAR
CASE eReqStatus OF
	E_CIP_Usage.eLocal:;
				eReqStatusLocal	:=E_CIP_Client_Selector.eClose;
	E_CIP_Usage.eTank_1,
	E_CIP_Usage.eTank_2:;
				eReqStatusLocal	:=E_CIP_Client_Selector.eMarinade_Up;	
	E_CIP_Usage.eTank_3,
	E_CIP_Usage.eTank_4:;
				eReqStatusLocal	:=E_CIP_Client_Selector.eColor_Up;	
	E_CIP_Usage.eTriBlender_Marinada,
	E_CIP_Usage.eLine_Marinada:;
				eReqStatusLocal	:=E_CIP_Client_Selector.eMarinade_Low;	
	E_CIP_Usage.eTriBlender_Color,
	E_CIP_Usage.eLine_Color:;
				eReqStatusLocal	:=E_CIP_Client_Selector.eColor_Low;	
	
END_CASE

IF eStatus=eReqStatusLocal 
AND eProcess=E_CIP_Client_Selector.eNone
AND eReq=E_CIP_Client_Selector.eNone
AND bReady
AND bDone
AND NOT bRun
THEN;
	m_CheckStatus:=TRUE;
END_IF
END_METHOD

METHOD m_Request_Reset : BOOL
VAR_IN_OUT
	memo: R_TRIG;
END_VAR
memo(CLK:=eReq=0);
IF TRUE 
AND memo.Q
THEN;
	SFCReset:=TRUE;
END_IF
END_METHOD

METHOD m_Run : BOOL
VAR_INPUT
	eReqProc			: E_CIP_Usage;
END_VAR
VAR
	eReqStatusLocal	: E_CIP_Client_Selector;
END_VAR
CASE eReqProc OF
	E_CIP_Usage.eLocal:;
				eReqStatusLocal	:=E_CIP_Client_Selector.eClose;
	E_CIP_Usage.eTank_1,
	E_CIP_Usage.eTank_2:;
				eReqStatusLocal	:=E_CIP_Client_Selector.eMarinade_Up;	
	E_CIP_Usage.eTank_3,
	E_CIP_Usage.eTank_4:;
				eReqStatusLocal	:=E_CIP_Client_Selector.eColor_Up;	
	E_CIP_Usage.eTriBlender_Marinada,
	E_CIP_Usage.eLine_Marinada:;
				eReqStatusLocal	:=E_CIP_Client_Selector.eMarinade_Low;	
	E_CIP_Usage.eTriBlender_Color,
	E_CIP_Usage.eLine_Color:;
				eReqStatusLocal	:=E_CIP_Client_Selector.eColor_Low;	
	
END_CASE

IF eProcess=E_CIP_Client_Selector.eNone THEN;
	eProcess:=eReq:=eReqStatusLocal;
	bDone:=FALSE;
	m_Run:=TRUE;
END_IF
END_METHOD

METHOD m_Set_SFCFlags_Reference : BOOL
//Set reference to SFC flags

refSFC.SFCInit REF= SFCInit;
refSFC.SFCReset REF= SFCReset;
refSFC.SFCError REF= SFCError;
refSFC.SFCEnableLimit REF= SFCEnableLimit;
refSFC.SFCErrorStep REF= SFCErrorStep;
refSFC.SFCErrorPOU REF= SFCErrorPOU;
refSFC.SFCQuitError REF= SFCQuitError;
refSFC.SFCPause REF= SFCPause;
refSFC.SFCTrans REF= SFCTrans;
refSFC.SFCCurrentStep REF= SFCCurrentStep;
refSFC.SFCTip REF= SFCTip;
refSFC.SFCTipMode REF= SFCTipMode;

// Cycle handle for SFC
m_SFC_Handle();
END_METHOD

END_FUNCTION_BLOCK

// ---- 03 Project/23 CIP/FB_CIP.TcPOU
FUNCTION_BLOCK FB_CIP EXTENDS FB_SFC_Cycle IMPLEMENTS ITF_FB_SFC_Cycle
VAR_INPUT
	valFillWater_T91	: E_Pis_Name;
	valFillWater_T92	: E_Pis_Name;
	valFillWater_T93	: E_Pis_Name;
	valFillWater_T94	: E_Pis_Name;
	
	lvlTank_T91			: ST_Tank_Level	;
	lvlTank_T92			: ST_Tank_Level	;
	lvlTank_T93			: ST_Tank_Level	;
	lvlTank_T94			: ST_Tank_Level	;

END_VAR
VAR_OUTPUT
END_VAR
VAR
	//bRun: BOOL;
	eRun: E_CIP_Source;

	eMode			: E_CIP_Mode;
	eCIP_Return		: E_CIP_Return;
	eCIP_Source		: E_CIP_Source;
	eCIP_Usage		: E_CIP_Usage;
	eReq			: ST_CIP_Request;
	eReqBlank		: ST_CIP_Request;
	eReqLocal		: ST_CIP_Request;
	
	ref_lvlTank_Client		: REFERENCE TO ST_Tank_Level	;

	//bStepDone: BOOL;
	
	iPosSelect_HMI: INT;

	rtPosMoveHMI_Up		: R_TRIG;
	rtPosMoveHMI_Down	: R_TRIG;
	rtPosDeleteHMI		: R_TRIG;
	rtPosDeleteAllHMI	: R_TRIG;
	
	eRefClient_fbElement		: REFERENCE TO FB_Element; // FB_Element // E_Element_State_Long
	bClientRef_done				: BOOL;
	fbElement_Blank				: FB_Element;
	eState_Long_Blank			: E_Element_State_Long;
	
	fbPis						: FB_Piston;
	stPis_FillWater_T91			: REFERENCE TO ST_Piston;
	stPis_FillWater_T92			: REFERENCE TO ST_Piston;
	stPis_FillWater_T93			: REFERENCE TO ST_Piston;
	stPis_FillWater_T94			: REFERENCE TO ST_Piston;
	
	rtReqLocalCIP_Full_HMI: R_TRIG;
	rtReqLocalCIP_Detergent_HMI: R_TRIG;
	rtReqCleanEmpty_HMI: R_TRIG;
	rtModeOff: R_TRIG;
	rtModeManual: R_TRIG;
	rtModeAuto: R_TRIG;
	bTemp: BOOL;
		
	//Process Control
	//concentration
	stDetergent					:	REFERENCE TO ST_ProcessControl	;
	pcDetergent					: 	REFERENCE TO FB_ProcessControl	;	//detergent local
	stDisInfectant				:	REFERENCE TO ST_ProcessControl	;
	pcDisInfectant				: 	REFERENCE TO FB_ProcessControl	;	//detergent local
    //temperature
	stHeatExchanger					:	REFERENCE TO ST_ProcessControl	;
	pcHeatExchanger					: 	REFERENCE TO FB_ProcessControl	;	//	
	stTemperature_Deterg			:	REFERENCE TO ST_ProcessControl	;
	pcTemperature_Deterg			: 	REFERENCE TO FB_ProcessControl	;	//detergent Client	
	stTemperature_Dis				:	REFERENCE TO ST_ProcessControl	;
	pcTemperature_Dis				: 	REFERENCE TO FB_ProcessControl	;//disinfectant local/client
	//temperature client return
	stTemp_ClntReturn				:	REFERENCE TO ST_ProcessControl	;//Client return temperature
	pcTemp_ClntReturn				: 	REFERENCE TO FB_ProcessControl	;//Client return temperature
	
	//flow rate
	stFlow1_Rate					:	REFERENCE TO ST_ProcessControl	;//CIP
	pcFlow1_Rate					: 	REFERENCE TO FB_ProcessControl	;//disinfectant local/client
	stFlow2_Rate					:	REFERENCE TO ST_ProcessControl	;//CIP send
	pcFlow2_Rate					: 	REFERENCE TO FB_ProcessControl	;//disinfectant local/client	return 
	stFlow3_Rate					:	REFERENCE TO ST_ProcessControl	;//CIP send
	pcFlow3_Rate					: 	REFERENCE TO FB_ProcessControl	;//disinfectant local/client	return 
	
	stColor_Level					:	REFERENCE TO ST_ProcessControl	;//CLient CIP //level control 
	pcColor_Level					: 	REFERENCE TO FB_ProcessControl	;//disinfectant local/client //level control 
	stMarinada_Level				:	REFERENCE TO ST_ProcessControl	;//CLient CIP //level control 
	pcMarinada_Level				: 	REFERENCE TO FB_ProcessControl	;//disinfectant local/client //level control 
	
	
